// calculate equatorial coordinates (used by Slew command, takes Alt/Az -> moves telescope)
fbHor2Eq(alt := fElevation, 
		az := fAzimuth,
		jd := fJd+fTimeOffset,
		lat := telescopeConfig.latitude,
		lon := telescopeConfig.longitude,
		altitude := telescopeConfig.altitude,
		alt_is_observed := FALSE,
		ra => fRightAscensionCalc,
		dec => fDeclinationCalc,
		ha => fHourAngleCalc);		
// caluclate pointing offsets
fbPointingForward(
	HourAngle	:= fHourAngleApparent,
	Declination	:= fDeclinationApparent,
	Latitude	:= telescopeConfig.latitude,
	HourAngle_correction => fHourAnglePointingOffset,
	Declination_correction => fDeclinationPointingOffset,
	HourAngle_velocity => fHourAngleVelocity,
	Declination_velocity => fDeclinationVelocity,
);
(*--------------------------------------------------------------*)
// get current coordinates (of motors)
fDeclinationCurrent := fbDeclination.ActualPosition ;
fHourAngleCurrent := fbHourAngle.ActualPosition ;
// calculte pointing inversion
fbPointingInversion(
	HourAngle:= fHourAngleCurrent,
	Declination:= fDeclinationCurrent,
	Latitude:=telescopeConfig.latitude,
	HourAngle_correction => fHourAngleInversionOffsetCalc,
	Declination_correction => fDeclinationInversionOffsetCalc,
	bValid => bPointingInversionValid
);
// near the horizon the inversion is chaotic and does not converge (see FB_PointingModelInversion);
// keep reporting the last trustworthy correction rather than whatever garbage it would return
IF bPointingInversionValid THEN
	fHourAngleInversionOffset := fHourAngleInversionOffsetCalc;
	fDeclinationInversionOffset := fDeclinationInversionOffsetCalc;
END_IF
(*--------------------------------------------------------------*)
// transform from apparent to icrs

//current
fbHaDec2RaDec(
	ha := fHourAngleCurrent,
	dec := fDeclinationCurrent,
	jd := fJd+fTimeOffset,
	lon := telescopeConfig.longitude,
	ra_out => fRightAscensionCurrentICRS,
	dec_out => fDeclinationCurrentICRS);
//current corrected
fbHaDec2RaDec(
	ha := fHourAngleCurrent - fHourAngleInversionOffset - F_HourAngleOffsetOnAxis(fHourAngleOffset, fDeclinationApparent),
	dec := fDeclinationCurrent - fDeclinationInversionOffset- fDeclinationOffset,
	jd := fJd+fTimeOffset,
	lon := telescopeConfig.longitude,
	ra_out => fRightAscensionCurrentICRScorr,
	dec_out => fDeclinationCurrentICRScorr);
(*--------------------------------------------------------------*)
// to ALT AZ
fbEq2Hor(
	ra := fRightAscensionCurrentICRS,
	dec := fDeclinationCurrentICRS,
	lon := telescopeConfig.longitude,
	lat := telescopeConfig.latitude,
	altitude := telescopeConfig.altitude,
	refract_to_observed := FALSE,
	JD := fJd + fTimeOffset,
	alt => fElevationCurrent,
	az => fAzimuthCurrent);
	
fbEq2Hor(
	ra := fRightAscensionCurrentICRScorr,
	dec := fDeclinationCurrentICRScorr,
	lon := telescopeConfig.longitude,
	lat := telescopeConfig.latitude,
	altitude := telescopeConfig.altitude,
	refract_to_observed := FALSE,
	JD := fJd + fTimeOffset,
	alt => fElevationCurrentSky,
	az => fAzimuthCurrentSky);
END_METHOD

// Hook of the template body (BROTLib#25 step 5.4, S3: the body of this block is the template text, the differences are in these methods). Horizon and pole-zone guards, limit homes, target checks.
METHOD PROTECTED _Guards
// #161: while an axis is uncalibrated (e.g. after a PLC activation) its counter is meaningless, so the horizon and
// pole-zone stops must not act on it, otherwise the power-on sweep and the jog are stopped. Protection then is the NC
// software limits, the sweep's DistanceLimit and the operator.
bAxesCalibrated := fbHourAngle.Calibrated AND fbDeclination.Calibrated;
// losing the reference while enabled and not homing: stop instead of silently releasing the horizon protection
rtrigCalibLost(CLK := bAxesCalibrated);
IF rtrigCalibLost.Q AND bReady AND NOT bError AND NOT aAxis[1].bHoming AND NOT aAxis[2].bHoming THEN
	_AutoStop();
END_IF
// #166: a running power-on does not move a calibrated axis, but enabling it is not settled for a few scans and the mount
// is not ready before stage 100, so a mount inside a limit was stopped and the power-on aborted (any bStop aborts it).
// Skip the automatic stop only while the axes that matter stand still; stage 100 hands over to bGoHome. Any motion, a
// user stop or an error still stops.
bPowerOnHold := bPowerActive AND NOT bError;
bHaMoving := aAxis[1].bInMotion OR aAxis[1].bInRamp OR aAxis[1].bHoming;
bDecMoving := aAxis[2].bInMotion OR aAxis[2].bInRamp OR aAxis[2].bHoming;
// If the Telescope dips under the fHorizon (e.g. while tracking, stop and gohome)
// (also gated on fPointingSafeAltitude so tracking never lingers in the pointing model's chaotic zone)
// #84: a park requested in a limit homes out of it first and then parks. The stop conditions are unchanged.
IF NOT bGoHomeActive THEN
	bLimitHome := FALSE;
END_IF
IF NOT bParkActive THEN
	bParkAfterHome := FALSE;
	bParkHomeDone := FALSE;
	bParkForceInPlace := FALSE;
END_IF
bInHorizonLimit := bAxesCalibrated AND fElevationCurrent < MAX(fHorizon+0.2, fPointingSafeAltitude);
bInPoleLimit := (fbDeclination.Calibrated AND fDeclinationCurrent > (90.0 - fPoleZone)) OR (bAxesCalibrated AND bTrackActive AND (fDeclinationApparent + fDeclinationOffset + fDeclinationPointingOffset > (90.0 - fPoleZone)));
IF bInHorizonLimit THEN
	IF NOT bSettled AND NOT bGoHomeActive AND NOT (bPowerOnHold AND NOT bHaMoving AND NOT bDecMoving) THEN
		_AutoStop();
	ELSIF bReady AND NOT bError AND NOT bParkHomeDone THEN	// #82: only when the home can run; the power-on homes (stage 100)
		bGoHomeActive := TRUE;
		bLimitHome := TRUE;		// #84: also when bGoHome was set already (Home(), power-on stage 100)
	END_IF
END_IF
// If the Telescope goes into the forbidden polezone (e.g. while tracking, stop and gohome)
IF bInPoleLimit THEN
	IF NOT bSettled AND NOT bGoHomeActive AND NOT (bPowerOnHold AND NOT bDecMoving) THEN
		_AutoStop();
	ELSIF bReady AND NOT bError AND NOT bParkHomeDone THEN	// #82: only when the home can run; the power-on homes (stage 100)
		bGoHomeActive := TRUE;
		bLimitHome := TRUE;		// #84
	END_IF
END_IF
//----------------------------------------------------------------------------------------------
// if the given coordinates to goto/slew are under the horizon
// (also rejects targets below fPointingSafeAltitude, where the pointing model's inversion is chaotic -- see FB_PointingModelInversion)
IF (bGotoActive AND (fElevationCalc < MAX(fHorizon + 1.0, fPointingSafeAltitude))) OR (bSlewActive AND (fElevation < MAX(fHorizon, fPointingSafeAltitude))) THEN
	// trigger event
	rtrigHorizonError(CLK:=TRUE);
	// reset input coords to parking position (always over horizon to stop bHorizonError from occuring)
	fDeclination := telescopeConfig.declinationPark;
	fbHaDec2RaDec(	jd := fJd +fTimeOffset,
					ha := telescopeConfig.houranglePark,
					dec := telescopeConfig.declinationPark,
					lon := telescopeConfig.longitude,
					ra_out => fRightAscension);
	// reset elevation values to abitrarry value over horizon, will get overwritten down the line
	fElevationCalc := 20.0;
	fElevation := 20.0;
	// stop telescope
	_AutoStop();
ELSE
	// reset event trigger
	rtrigHorizonError(CLK:=FALSE);
END_IF

// if the given coordinates to goto/slew are in the PoleZone
IF (bGotoActive AND (fDeclinationApparent > (90.0 - fPoleZone))) OR (bSlewActive AND (fDeclinationCalc  > (90.0 - fPoleZone))) THEN
	// trigger event
	rtrigPoleError(CLK:=TRUE);
	// reset input coords to parking position (always over horizon to stop bHorizonError from occuring)
	fDeclination := telescopeConfig.declinationPark;
	fbHaDec2RaDec(	jd := fJd +fTimeOffset,
					ha := telescopeConfig.houranglePark,
					dec := telescopeConfig.declinationPark,
					lon := telescopeConfig.longitude,
					ra_out => fRightAscension);
	// reset elevation values to abitrarry value over horizon, will get overwritten down the line
	fElevationCalc := 20.0;
	fElevation := 20.0;
	// stop telescope
	_AutoStop();

ELSE
	// reset event trigger
	rtrigPoleError(CLK:=FALSE);
END_IF
END_METHOD

// Hook of the template body (BROTLib#25 step 5.4, S3: the body of this block is the template text, the differences are in these methods). Power-on warning, idle park, state-machine timeouts, pending home and park.
METHOD PROTECTED _Timers
tpPowerOnWarning(IN := bPowerActive OR (NOT fbHourAngle.bEnable), PT := T#250MS);

tonPowerTimeout(IN := TCS_command = E_TCSCommand.no_command AND NOT bIsParked, PT := T#12H, nDivisor := nTimeDivisor);
// MONETcommon#17: state-machine timeouts, checked in _GotoTelescope/_HomeTelescope/_SlewTelescope
// #75: count only while the command is the one being run (TCS_command is last scan's dispatch) and without an error.
// Counting from the request, a command that never started (not ready, preempted) fired the timeout in the next
// stop/park/reset after 600 s and latched an error, and with the horizon/pole auto-home setting bGoHome again every
// scan the timer never dropped, so no reset cleared it.
tonGotoTimeout(IN := bGotoActive AND TCS_command = E_TCSCommand.goto AND NOT bError, PT := T#600S, nDivisor := nTimeDivisor);
tonHomeTimeout(IN := bGoHomeActive AND TCS_command = E_TCSCommand.gohome AND NOT bError, PT := T#600S, nDivisor := nTimeDivisor);
tonSlewTimeout(IN := bSlewActive AND TCS_command = E_TCSCommand.slew AND NOT bError, PT := T#600S, nDivisor := nTimeDivisor);
tonParkTimeout(IN := bParkActive AND TCS_command = E_TCSCommand.park AND NOT bError, PT := T#600S, nDivisor := nTimeDivisor);
// #75: a Home() that never starts (axes off, telescope not ready) left bGoHome set for good, swallowing Track() and
// Slew(). Drop it after 2 min, with a log line, without an error. Not at once: the home that the power-on requests in
// stage 100 can wait a few scans for bReady, and a stop from slew speed takes about 4 s. Not during a power-on.
tonHomePending(IN := bGoHomeActive AND TCS_command <> E_TCSCommand.gohome AND NOT bPowerActive AND NOT bError, PT := T#2M, nDivisor := nTimeDivisor);
IF tonHomePending.Q THEN
    fbStartup.MarkAbortedIfInitializing();
	bGoHomeActive := FALSE;
	// #108: say what was pending. "Not ready, power on" was also logged when a stop before the home had not finished.
	fbHomeDrop(bReady := bReady, bStopPending := TCS_command = E_TCSCommand.stop OR NOT bSettled);
	sHomeEnd := fbHomeDrop.sEnd;
	sHomeDropWhy := fbHomeDrop.sWhy;
	bHomeCancelled := TRUE;
END_IF
// #197: a park that is requested but not started (not dispatched, not in the axes-off path, no stop or home running)
// waited without a timeout: tonParkTimeout counts only a running park (#75). After 2 min: say why and park in place.
tonParkPending(IN := bParkActive AND TCS_command <> E_TCSCommand.park AND TCS_command <> E_TCSCommand.gohome
	AND NOT bMoveAbortPending AND NOT bError AND NOT bEstopTriggered AND NOT bParkForceInPlace, PT := T#2M, nDivisor := nTimeDivisor);
IF tonParkPending.Q THEN
	bParkForceInPlace := TRUE;
	fbHomeDrop(bReady := bReady, bStopPending := TCS_command = E_TCSCommand.stop OR NOT bSettled);
	TCSparkErrorEvent.OnMessage := CONCAT(CONCAT('Park did not start within 2 min (', fbHomeDrop.sWhy), '): parking in place with the axes off.');
	bParkInError := TRUE;
END_IF
IF tonPowerTimeout.Q AND NOT bIsParked THEN
	bParkActive := TRUE;
	// #83: fire once. With the axes off or in error the park does not set bIsParked, so Q stayed TRUE and bPark was
	// set again every scan (dropping Track/Goto/Slew/Home, re-commanding the dome). The timer counts again from now.
	tonPowerTimeout(IN := FALSE);
END_IF
END_METHOD

// Hook of the template body (BROTLib#25 step 5.4, S3: the body of this block is the template text, the differences are in these methods). The replacement gets its own timeout.
METHOD PROTECTED _RestartMoveTimeout
VAR_INPUT
	eKeep	: E_TCSCommand;
END_VAR
CASE eKeep OF
	E_TCSCommand.gohome:	tonHomeTimeout(IN := FALSE, PT := T#600S, nDivisor := nTimeDivisor);
	E_TCSCommand.goto:		tonGotoTimeout(IN := FALSE, PT := T#600S, nDivisor := nTimeDivisor);
	E_TCSCommand.slew:		tonSlewTimeout(IN := FALSE, PT := T#600S, nDivisor := nTimeDivisor);
END_CASE
END_METHOD

// Hook of the template body (BROTLib#25 step 5.4, S3: the body of this block is the template text, the differences are in these methods). The automatic parks.
METHOD PROTECTED _ParkRequests
// BROTLib#25 step 4.4d (decided by Tim 2026-11-09: MONETcommon wins): a new hardware error (hour angle, declination or focus; not a
// software or cabinet error) while not parked and without E-stop starts the park by itself, like MONETcommon#86. The park branch
// below does what is safe without the mount (the axes are disabled by the error): covers close, dome parks, focus off; the mount
// is not moved and bIsParked is not set until the covers are closed and the dome is parked. A running power-on is aborted by
// the park (#109). Edge only: a still present error does not start it again.
bErrorParkStarted := BROTLib.F_ErrorParkRequest(
	bHwError := fbHourAngle.Error OR fbDeclination.Error OR (fbFocus <> 0 AND_THEN fbFocus.Error),
	bHwErrorLast := bHwErrorLast,
	bIsParked := bIsParked,
	bEstop := bEstopTriggered);
bHwErrorLast := fbHourAngle.Error OR fbDeclination.Error OR (fbFocus <> 0 AND_THEN fbFocus.Error);
IF bErrorParkStarted THEN
	Park();
END_IF
END_METHOD

// Hook of the template body (BROTLib#25 step 5.4, S3: the body of this block is the template text, the differences are in these methods). TRUE: the pending park waits. The gate (no stop, no power-on, no abort stop) is in the body.
METHOD PROTECTED _ParkPreStep : BOOL
_ParkPreStep := FALSE;
bTrackActive := FALSE;
IF bError OR bEstopTriggered OR (TCS_command <> E_TCSCommand.park AND NOT fbHourAngle.Enable AND NOT fbDeclination.Enable) THEN
	_ParkInPlace();
	_ParkPreStep := TRUE;
ELSIF (NOT bIsPowered OR bParkForceInPlace) AND TCS_command <> E_TCSCommand.park THEN
	// #197: no completed power-on (aborted by this park, or stopped in stage 40 or later) but an axis is on: the park can
	// never be dispatched. Switch the axes off once they are at rest, then the axes-off park parks in place.
	// TCS_command must not stay on poweron: _PowerOn and its 12 h timeout would stay selected.
	fbSweepStop.ArmAll();
	TCS_command := E_TCSCommand.no_command;
	_ParkPreStep := TRUE;
ELSIF bGoHomeActive AND bLimitHome THEN
	// #84: a park in a limit: the home out of the limit runs first (the arbiter dispatches it), the park follows (bParkHomeDone)
	IF NOT bParkAfterHome THEN
		bParkAfterHome := TRUE;
		bParkHomeFirst := TRUE;
	END_IF
	_ParkPreStep := TRUE;
ELSIF NOT (bReady AND NOT bBusy) THEN
	_ParkPreStep := TRUE;
END_IF
END_METHOD

// Hook of the template body (BROTLib#25 step 5.4, S3: the body of this block is the template text, the differences are in these methods). The arbiter input bEmergencyPark.
METHOD PROTECTED _EmergencyPark : BOOL
_EmergencyPark := FALSE;
END_METHOD

// Hook of the template body (BROTLib#25 step 5.4, S3: the body of this block is the template text, the differences are in these methods). The arbiter input bStopped: at rest and no stop transaction running.
METHOD PROTECTED _AtRest : BOOL
_AtRest := bSettled;	// IAG50cm: at rest and no stop transaction running
END_METHOD

// Hook of the template body (BROTLib#25 step 5.4, S3: the body of this block is the template text, the differences are in these methods). The arbiter interrupts the power-on.
METHOD PROTECTED _InterruptPower
IF _PowerOnStage() >= 40 THEN	// abort path: bPowerActive FALSE, startup marked aborted, stage 0; returns the stage it was in
	IF fbArbiter.bPowerAbortedByPark THEN
		// #197: the axes are on and may be sweeping: stop them. The park then switches them off (nothing else can: bReady
		// needs the completed power-on) and parks in place.
		fbSweepStop.ArmAll();
	ELSE
		fbSweepStop.Arm();		// #113: stopped in the calibration sweep (stage 40 and later)
	END_IF
	fbHourAngle.bStopSweep := TRUE;		// #198: no new sweep step after this stop, also before the sweep has started
	fbDeclination.bStopSweep := TRUE;
END_IF
END_METHOD

// Hook of the template body (BROTLib#25 step 5.4, S3: the body of this block is the template text, the differences are in these methods). The arbiter interrupts the park.
METHOD PROTECTED _InterruptPark
IF bWasPark THEN
	sParkEnd := 'cancelled by stop';
	fbSweepStop.Cancel();		// #197: the park is gone, the axes stay as they are
END_IF
_DoPark();
END_METHOD

// Hook of the template body (BROTLib#25 step 5.4, S3: the body of this block is the template text, the differences are in these methods). The arbiter interrupts the goto.
METHOD PROTECTED _InterruptGoto
_DoGoto();
END_METHOD

// Hook of the template body (BROTLib#25 step 5.4, S3: the body of this block is the template text, the differences are in these methods). The arbiter interrupts the slew.
METHOD PROTECTED _InterruptSlew
_DoSlew();
END_METHOD

// Hook of the template body (BROTLib#25 step 5.4, S3: the body of this block is the template text, the differences are in these methods). The arbiter interrupts the home.
METHOD PROTECTED _InterruptGoHome
IF bWasGoHome THEN
	IF bStopActive THEN
		sHomeEnd := 'cancelled by stop';	// #84: also the home that a park waited for
	ELSE
		sHomeEnd := 'cancelled by park';
	END_IF
END_IF
_DoGoHome();
END_METHOD

// Hook of the template body (BROTLib#25 step 5.4, S3: the body of this block is the template text, the differences are in these methods). After the arbiter has been applied.
METHOD PROTECTED _AfterArbiter
// #196: the axes are off, there is nothing to stop; the covers have no stop command and the park goes on
IF bStopActive AND bSafeParked AND NOT bWasPark AND NOT bWasPower AND NOT bWasMove AND NOT bWasGoHome THEN
	bStopIgnored := TRUE;
END_IF
END_METHOD

// Hook of the template body (BROTLib#25 step 5.4, S3: the body of this block is the template text, the differences are in these methods). Idle: the axis commands are dropped.
METHOD PROTECTED _DropAxisCommands
	fbHourAngle.MoveAxis := FALSE;
	fbDeclination.MoveAxis := FALSE;
	fbHourAngle.bTracking := FALSE;
	fbDeclination.bTracking := FALSE;
END_METHOD

// Hook of the template body (BROTLib#25 step 5.4, S3: the body of this block is the template text, the differences are in these methods). TCS_command changed.
METHOD PROTECTED _OnCommandChanged
// #108: a stop transaction starts here and lasts as long as TCS_command stays stop (also through the wait of a
// gohome that preempted a track): each axis gets one stop in it
IF TCS_command = E_TCSCommand.stop THEN
	fbStopTx.Begin();
END_IF
END_METHOD

// Calls the stage machine of the power-on; returns the stage it was in (>= 40: the sweep stop of the power-on runs).
METHOD PRIVATE _PowerOnStage : USINT
_PowerOnStage := _PowerOn();
END_METHOD

// Hook of the template body (BROTLib#25 step 5.4). Calls the stage machine of the power-on.
METHOD PROTECTED _DoPowerOn
_PowerOnStage();
END_METHOD

// Hook of the template body (BROTLib#25 step 5.4, S3: the body of this block is the template text, the differences are in these methods). Calls the stage machine.
METHOD PROTECTED _DoPark
_ParkTelescope();
END_METHOD

// Hook of the template body (BROTLib#25 step 5.4, S3: the body of this block is the template text, the differences are in these methods). Calls the stage machine.
METHOD PROTECTED _DoGoHome
_HomeTelescope();
END_METHOD

// Hook of the template body (BROTLib#25 step 5.4, S3: the body of this block is the template text, the differences are in these methods). Calls the stage machine.
METHOD PROTECTED _DoGoto
_GotoTelescope();
END_METHOD

// Hook of the template body (BROTLib#25 step 5.4, S3: the body of this block is the template text, the differences are in these methods). Calls the stage machine.
METHOD PROTECTED _DoSlew
_SlewTelescope();
END_METHOD

// Hook of the template body (BROTLib#25 step 5.4, S3: the body of this block is the template text, the differences are in these methods). Calls the stage machine.
METHOD PROTECTED _DoTrack
_TrackTelescope();
END_METHOD

// Hook of the template body (BROTLib#25 step 5.4, S3: the body of this block is the template text, the differences are in these methods). Calls the stage machine.
METHOD PROTECTED _DoStop
_StopTelescope();
END_METHOD

// Hook of the template body (BROTLib#25 step 5.4, S3: the body of this block is the template text, the differences are in these methods). The timeout of a command.
METHOD PROTECTED _CommandTimeout : TIME
VAR_INPUT
	eCommand	: E_TCSCommand;
END_VAR
CASE eCommand OF
	E_TCSCommand.poweron:	_CommandTimeout := T#12H;
	E_TCSCommand.stop:		_CommandTimeout := T#30S;	// #40: a stop from slew speed takes about 4 s, a preempting stop can follow a long move
	E_TCSCommand.track:		_CommandTimeout := T#12H;
ELSE
	_CommandTimeout := T#2M;
END_CASE
END_METHOD

// Hook of the template body (BROTLib#25 step 5.4, S3: the body of this block is the template text, the differences are in these methods). After the dispatch.
METHOD PROTECTED _AfterDispatch
// nothing
END_METHOD

// Hook of the template body (BROTLib#25 step 5.4, S3: the body of this block is the template text, the differences are in these methods). Motion, stop transaction, sweep stop, readiness and the in-place park status.
METHOD PROTECTED _UpdateStatus
(* STATUS BOOLS*)
bSliding := NOT bTracking AND (aAxis[1].bInMotion OR aAxis[1].bInRamp OR
			aAxis[2].bInMotion OR aAxis[2].bInRamp );

// signal must be stable for 1s
tonTrackingDelay(in := aAxis[1].bTracking AND
			aAxis[2].bTracking ,PT :=T#1000MS, Q => bTracking);

// #92: a move that was commanded (MoveAxis -> MoveTo) is reported by the NC a few cycles later; until then the axis
// reports StandStill. A stop in that window saw bStopped, so bStop was cleared after one scan, the stop only dropped
// MoveAxis (which does not cancel a move that has started) and no axis stop was sent: the move ran to its end (T18.4,
// park, Dec). The axis is not at rest while its move is on the way; the stop then lasts until the axis moves and gets
// its axis stop from the stop transaction.
rtHaMove(CLK := fbHourAngle.MoveAxis);
rtDecMove(CLK := fbDeclination.MoveAxis);
IF rtHaMove.Q THEN
	bHaMovePending := TRUE;
END_IF
IF rtDecMove.Q THEN
	bDecMovePending := TRUE;
END_IF
IF aAxis[1].bInMotion OR aAxis[1].bInRamp OR aAxis[1].bHoming OR fbHourAngle.MoveDone OR bError OR NOT fbHourAngle.bEnable THEN
	bHaMovePending := FALSE;
END_IF
IF aAxis[2].bInMotion OR aAxis[2].bInRamp OR aAxis[2].bHoming OR fbDeclination.MoveDone OR bError OR NOT fbDeclination.bEnable THEN
	bDecMovePending := FALSE;
END_IF
tonHaMovePending(IN := bHaMovePending, PT := T#1S);
tonDecMovePending(IN := bDecMovePending, PT := T#1S);
IF tonHaMovePending.Q THEN
	bHaMovePending := FALSE;
END_IF
IF tonDecMovePending.Q THEN
	bDecMovePending := FALSE;
END_IF

// #198: a pause of the calibration sweep reports StandStill, but FB_LatchHome is still in its sequence (or about to start
// it): the axis is not at rest. A stop in a pause saw bStopped, ran for one scan and sent no axis stop.
bStopped :=  (NOT fbHourAngle.bEnable OR (aAxis[1].bStandStill AND NOT fbHourAngle.bSweepActive)) AND
			(NOT fbDeclination.bEnable OR (aAxis[2].bStandStill AND NOT fbDeclination.bSweepActive)) AND
			NOT bHaMovePending AND NOT bDecMovePending;

// #98: bStopped is TRUE for one scan at the start of every stop, before MC_Stop has taken hold (StandStill is still
// TRUE), and a home commanded while MC_Stop locks the axis (StateDWord bit 29) fails with 17135. A stop transaction
// is settled when every axis that was sent a stop reported Done and no axis has been locked for 3 scans.
IF bResetActive OR bError OR bEstopTriggered THEN
	fbStopTx.Cancel();
	fbSweepStop.Cancel();
END_IF
_SetStopTxInputs();
fbStopTx.Monitor();
bSettled := bStopped AND NOT fbStopTx.bActive;

// #120: a stop transaction that is not settled 30 s after it began (an axis never reported Done) no longer waits for the
// Done: it settles as soon as the telescope is at rest. The stop is not sent again. Clear StopAxis of the axes without a
// Done so that the next stop gives a rising edge (FB_AxisControl.StopAxis) and the home hold does not see a stale stop.
IF fbStopTx.bTimedOut THEN
	IF fbStopTx.abNoDone[1] AND fbStopTx.abNoDone[2] THEN
		sStopNoDone := 'HA and Dec';
	ELSIF fbStopTx.abNoDone[1] THEN
		sStopNoDone := 'HA';
	ELSE
		sStopNoDone := 'Dec';
	END_IF
	IF NOT fbStopTx.bActive THEN
		TCSstopTimeoutEvent.OnMessage := CONCAT(CONCAT('STOP: no stop Done from ', sStopNoDone), ' within 30 s; telescope at rest, stop released.');
	ELSIF NOT bStopped THEN
		TCSstopTimeoutEvent.OnMessage := CONCAT(CONCAT('STOP: no stop Done from ', sStopNoDone), ' within 30 s; axes still moving, released when at rest.');
	ELSE
		TCSstopTimeoutEvent.OnMessage := CONCAT(CONCAT('STOP: no stop Done from ', sStopNoDone), ' within 30 s; axis locked (stop active) or homing, released when it ends.');
	END_IF
	bStopTimeoutLog := TRUE;
ELSIF fbStopTx.bForced THEN
	TCSstopTimeoutEvent.OnMessage := 'STOP released: at rest without a stop Done from an axis (30 s timeout).';
	bStopTimeoutLog := TRUE;
END_IF
IF fbStopTx.bForced THEN
	IF fbStopTx.abNoDone[1] THEN
		fbHourAngle.StopAxis := FALSE;
	END_IF
	IF fbStopTx.abNoDone[2] THEN
		fbDeclination.StopAxis := FALSE;
	END_IF
END_IF

// #113: a stop in the calibration sweep leaves the axes enabled and uncalibrated; once the stop has settled and the
// homing is aborted, switch the uncalibrated axes off (the next power-on starts the sweep again), READY_STATE -2
IF bPowerActive THEN
	fbSweepStop.Cancel();
END_IF
fbSweepStop(bSettled := bSettled,
			bHaCalibrated := fbHourAngle.bCalibrated, bDecCalibrated := fbDeclination.bCalibrated,
			bHaHoming := fbHourAngle.fbLatchHome.Busy, bDecHoming := fbDeclination.fbLatchHome.Busy,
			bOtherBusy := fbFocus <> 0 AND_THEN fbFocus.Busy);
IF fbSweepStop.bDisableHa THEN
	fbHourAngle.Enable := FALSE;
END_IF
IF fbSweepStop.bDisableDec THEN
	fbDeclination.Enable := FALSE;
END_IF
			
bHomed := fbHourAngle.bCalibrated AND fbDeclination.bCalibrated AND (fbFocus <> 0 AND_THEN fbFocus.Calibrated);
			
bReady := bHomed AND 
	bIsPowered AND 
	fbHourAngle.bEnable AND
	fbDeclination.bEnable AND
	(fbFocus <> 0 AND_THEN fbFocus.Enable) AND
    NOT bError;

bBusy := aAxis[1].bBusy OR aAxis[2].bBusy OR (fbFocus <> 0 AND_THEN fbFocus.Busy);
//----------------------------------------------------------------------------------------------
(* STATUS STATES*)
// Public completion is latched only by the final startup stage, never by mechanical bReady alone.
// #110: the covered state ends with a power-on, an error or an E-stop.
IF bSafeParked AND (bPowerActive OR bError OR bEstopTriggered) THEN
	// #200: every exit of the in-place park has an end line
	IF bEstopTriggered THEN
		sParkInPlaceEnd := 'aborted: E-stop pressed, the covers and the dome cannot move. Release it, reset, then park again.';
		nParkInPlaceLevel := ADSLOG_MSGTYPE_WARN;
	ELSIF bError THEN
		IF fbCovers.Closed THEN
			sParkInPlaceEnd := 'aborted by an error: covers closed, the mount was not moved. Reset, then park again.';
		ELSE
			sParkInPlaceEnd := 'aborted by an error: covers closing, the mount was not moved. Reset, then park again.';
		END_IF
		nParkInPlaceLevel := ADSLOG_MSGTYPE_WARN;
	ELSE
		sParkInPlaceEnd := 'cancelled by power-on';
		nParkInPlaceLevel := ADSLOG_MSGTYPE_HINT;
	END_IF
	bParkInPlaceDone := TRUE;
END_IF
IF bPowerActive OR bError OR bEstopTriggered THEN
    bSafeParked := FALSE;
END_IF
// #187: an axes-off park (power-on aborted by a park, park after a stopped power-on) ends parked, like a park of MONET:
// bIsParked means covers closed and dome parked with the axes off, bParkedInPlace says the mount was not moved.
// Without it bIsParked stayed FALSE, and the 12 h idle park fired again every 12 h.
tonParkInPlace(IN := bSafeParked AND NOT bIsParked, PT := T#120S, nDivisor := nTimeDivisor);
IF bSafeParked AND fbCovers.Closed AND fbDome.Parked THEN
	IF NOT bIsParked OR bParkInPlaceOpen THEN
		bIsParked := TRUE;
		bParkedInPlace := TRUE;
		sParkInPlaceEnd := 'completed in place: covers closed, dome parked, the mount stays where it stood (#187)';
		nParkInPlaceLevel := ADSLOG_MSGTYPE_HINT;
		bParkInPlaceDone := TRUE;
	END_IF
	bIsPowered := FALSE;
	bSafeParked := FALSE;
ELSIF bSafeParked AND (tonParkInPlace.Q OR fbDome.Error) THEN
	// give up: not 0.3 for ever. The park start line said what was requested; this is the end line (#200).
	bSafeParked := FALSE;
	sParkInPlaceEnd := 'aborted: the covers did not close or the dome did not park within 120 s, or the dome is in error.';
	nParkInPlaceLevel := ADSLOG_MSGTYPE_WARN;
	bParkInPlaceDone := TRUE;
END_IF
END_METHOD

// Hook of the template body (BROTLib#25 step 5.4, S3: the body of this block is the template text, the differences are in these methods). The Parking input of the READY_STATE.
METHOD PROTECTED _ReadyStateParking : BOOL
_ReadyStateParking := (bParkActive OR bSafeParked) AND NOT bPowerActive;
END_METHOD

// Hook of the template body (BROTLib#25 step 5.4, S3: the body of this block is the template text, the differences are in these methods). The slewing flag of the motion state.
METHOD PROTECTED _IsSlewing : BOOL
_IsSlewing := bSliding;
END_METHOD

// Hook of the template body (BROTLib#25 step 5.4, S3: the body of this block is the template text, the differences are in these methods). The stop transaction has settled.
METHOD PROTECTED _StopSettled : BOOL
_StopSettled := bSettled;
END_METHOD

// Hook of the template body (BROTLib#25 step 5.4, S3: the body of this block is the template text, the differences are in these methods). The abort stop has been released.
METHOD PROTECTED _OnAbortStopReleased
// nothing
END_METHOD

// Hook of the template body (BROTLib#25 step 5.4, S3: the body of this block is the template text, the differences are in these methods). The reset is released.
METHOD PROTECTED _ReleaseReset
// unset the RESET command when no Error is present
IF NOT bError THEN
	bResetActive := FALSE;
END_IF
END_METHOD

// Hook of the template body (BROTLib#25 step 5.4, S3: the body of this block is the template text, the differences are in these methods). End of the scan: the drives are cut on an E-stop.
METHOD PROTECTED _SafeStateEndOfScan
IF bEstopTriggered THEN
	fbHourAngle.Enable := FALSE;
	fbDeclination.Enable := FALSE;
END_IF
END_METHOD

// Hook of the template body (BROTLib#25 step 5.4, S3: the body of this block is the template text, the differences are in these methods). The period of the telemetry.
METHOD PROTECTED _TelemetryPeriod : TIME
IF bSliding OR bTrackActive OR bTracking THEN
	_TelemetryPeriod := T#1000MS;	// during movement every second
ELSE
	_TelemetryPeriod := T#5000MS;	// otherwise every five seconds
END_IF
END_METHOD

// Hook of the template body (BROTLib#25 step 5.4, S3: the body of this block is the template text, the differences are in these methods). Sends the telemetry.
METHOD PROTECTED _SendTelemetry : BOOL
THIS^._SendTelemetryEquitorial();
END_METHOD

// Hook of the template body (BROTLib#25 step 5.4, S3: the body of this block is the template text, the differences are in these methods). End of the scan.
METHOD PROTECTED _EndOfScan
IF NOT bGoHomeActive AND TCS_command <> E_TCSCommand.gohome THEN
	bHomeByCommand := FALSE;	// the commanded home is over
END_IF
END_METHOD

// plan step 3.4: the event function blocks at the end of the body (ADS log and MQTT log), moved unchanged; called at the end of the body.
METHOD PROTECTED _LogEvents
VAR_INPUT
END_VAR
(* Event function blocks start here. *)
TCSpowerEvent(	Trigger := bPowerFailure, 
				Level := ADSLOG_MSGTYPE_ERROR,
				FormatString := 'power %s',
				//OnMessage := 'Failure',
				OffMessage := 'OK', 
				Comm := fbComm);

TCSgohomeEvent.OffMessage := sHomeEnd;		// #75: "GOHOME completed" was also logged when the home was cancelled or timed out
TCSgohomeEvent(	Trigger := bGoHomeActive, 
				Level := ADSLOG_MSGTYPE_HINT,
				FormatString := 'GOHOME %s',
				OnMessage := 'commencing',
				Comm := fbComm);
sHomeEnd := 'completed';
// #197/#200: the in-place park that goes on from a logged park ends with the PARK end line, one per park
IF bParkInPlaceDone AND bParkInPlaceOpen THEN
	sParkEnd := sParkInPlaceEnd;
	TCSparkEvent.OffLevel := nParkInPlaceLevel;
	bParkInPlaceOpen := FALSE;
	bParkInPlaceDone := FALSE;
END_IF
TCSparkEvent.OffMessage := sParkEnd;		// #57: "PARK completed" was also logged when the park was cancelled
TCSparkEvent(	Trigger := bParkActive OR bParkInPlaceOpen,
				Level := ADSLOG_MSGTYPE_HINT,
				FormatString := 'PARK %s',
				OnMessage := 'commencing',
				Comm := fbComm);
TCSparkInPlaceEvent(	Trigger := bParkInPlaceDone,
				Level := nParkInPlaceLevel,
				FormatString := 'PARK %s',
				OnMessage := sParkInPlaceEnd,
				Comm := fbComm);
bParkInPlaceDone := FALSE;
bParkLogged := bParkActive;
sParkEnd := 'completed';
TCSparkEvent.OffLevel := ADSLOG_MSGTYPE_HINT;
TCSgotoEvent(	Trigger := bGotoActive, 
				Level := ADSLOG_MSGTYPE_HINT,
				FormatString := 'GOTO %s',
				OnMessage := 'commencing',
				OffMEssage := 'completed', 
				Comm := fbComm);
TCStrackEvent(	Trigger := bTrackActive, 
				Level := ADSLOG_MSGTYPE_HINT,
				FormatString := 'TRACK %s',
				OnMessage := 'commencing',
				OffMEssage := 'completed', 
				Comm := fbComm);
TCSstopEvent(	Trigger := bStopActive, 
				Level := ADSLOG_MSGTYPE_WARN,
				FormatString := 'STOP %s',
				OnMessage := 'commencing',
				OffMEssage := 'completed',
				OffLevel := ADSLOG_MSGTYPE_HINT, 
				Comm := fbComm);
TCSstopIgnoredEvent(	Trigger := bStopIgnored,
				Level := ADSLOG_MSGTYPE_WARN,
				FormatString := '%s',
				OnMessage := 'Stop ignored: the covers and the dome cannot be stopped, the in-place park continues.',
				Comm := fbComm);
bStopIgnored := FALSE;
TCStargetHorizonEvent(	Trigger := rtrigHorizonError.Q, 
				Level := ADSLOG_MSGTYPE_WARN,
				FormatString := '%s',
				OnMessage := 'Target below safe horizon, stopping telescope.',
				OffMEssage := '', 
				Comm := fbComm);
TCSaltitudeEvent(	Trigger := bAxesCalibrated AND fElevationCurrent<MAX(fHorizon+2.0, fPointingSafeAltitude+2.0),
				Level := ADSLOG_MSGTYPE_WARN,
				FormatString := '%s',
				OnMessage := 'Telescope below safe horizon, aboard and slew telescope to home position.',
				OffMEssage := '', 
				Comm := fbComm);
TCSnearPoleEvent(	Trigger := rtrigPoleError.Q, 
				Level := ADSLOG_MSGTYPE_WARN,
				FormatString := '%s',
				OnMessage := 'Target to close to the celestial pole, stopping telescope.',
				OffMEssage := '', 
				Comm := fbComm);			
TCSreadyEvent(	Trigger := bReady, 
				Level := ADSLOG_MSGTYPE_HINT,
				FormatString := '%s',
				OnMessage := 'IAG50cm startup finished', 
				Comm := fbComm);
TCSparkErrorEvent(	Trigger := bParkInError,
				Level := ADSLOG_MSGTYPE_WARN,
				FormatString := '%s',
				// OnMessage is set in the arbitration (texts built from sParkWhy); a literal here overwrote it (#57)
				Comm := fbComm);
bParkInError := FALSE;
TCShomeCancelEvent(	Trigger := bHomeCancelled,
				Level := ADSLOG_MSGTYPE_WARN,
				FormatString := '%s',
				OnMessage := CONCAT('Home request dropped: ', sHomeDropWhy),
				Comm := fbComm);
bHomeCancelled := FALSE;
TCSpowerBlockedEvent(	Trigger := bPowerBlocked,
				Level := ADSLOG_MSGTYPE_ERROR,
				FormatString := '%s',
				Comm := fbComm);
bPowerBlocked := FALSE;
TCSparkHomeEvent(	Trigger := bParkHomeFirst,
				Level := ADSLOG_MSGTYPE_HINT,
				FormatString := '%s',
				OnMessage := 'Park in the horizon/pole-zone limit: homing out of it first, then parking',
				Comm := fbComm);
bParkHomeFirst := FALSE;
TCSpowerParkEvent(	Trigger := bPowerAbortedByPark,
				Level := ADSLOG_MSGTYPE_WARN,
				FormatString := '%s',
				OnMessage := 'Power-on aborted by park',
				Comm := fbComm);
bPowerAbortedByPark := FALSE;
TCSinitRefusedEvent(	Trigger := bInitRefused,
				Level := ADSLOG_MSGTYPE_WARN,
				FormatString := 'power-on ignored: %s',
				OnMessage := sInitRefusedReason,
				Comm := fbComm);
bInitRefused := FALSE;
// every rejection is logged (ADS log and MQTT log topic); an identical one repeated within 2 s once, all are counted. The event is
// re-armed with FALSE first so that rejections in consecutive scans each give a rising edge (as MONETcommon).
tonRejectRepeat(IN := TRUE, PT := T#2S);
RejectEvent(Trigger := FALSE, Comm := fbComm);
IF bCommandRejected THEN
	IF tonRejectRepeat.Q OR eLastRejectedCommand <> eLoggedCommand OR eLastRejectReason <> eLoggedReason THEN
		sRejectMessage := CONCAT(CONCAT(BROTLib.F_TCSCommandText(eLastRejectedCommand), ' rejected: '),
			BROTLib.F_CommandRejectText(eLastRejectReason));
		RejectEvent(Trigger := TRUE, Level := ADSLOG_MSGTYPE_WARN, FormatString := '%s',
			OnMessage := sRejectMessage, Comm := fbComm);
		eLoggedCommand := eLastRejectedCommand;
		eLoggedReason := eLastRejectReason;
		tonRejectRepeat(IN := FALSE);
	END_IF
	bCommandRejected := FALSE;
END_IF
TCSstopTimeoutEvent(	Trigger := bStopTimeoutLog,
				Level := ADSLOG_MSGTYPE_WARN,
				FormatString := '%s',
				Comm := fbComm);
bStopTimeoutLog := FALSE;
TCSsoftErrorEvent(	Trigger := bSoftwareError,
				Level := ADSLOG_MSGTYPE_ERROR,
				FormatString := 'Command timeout error %s',	// 16 goto, 32 park, 48 gohome, 64 slew (16#10, 16#20, 16#30, 16#40)
				OnMessage := UDINT_TO_STRING(nSoftwareErrorID),
				OffMessage := 'reset',
				Comm := fbComm);
TCSCTOEvent(	Trigger := tonCommandTimeout.Q,
				Level := ADSLOG_MSGTYPE_WARN,
				FormatString := 'A timeout occured during %s command!',
				Comm := fbComm);
END_METHOD

// The state BROTLib.F_CommandAcceptance decides on. eExcludeOwn leaves the own request out of bMoveActive. bMoveAbortPending stands in for
// bMoveAbortPending until the abort stop (command model step 3A).
METHOD PRIVATE _CommandState : BROTLib.ST_CommandState
VAR_INPUT
	eExcludeOwn	: E_TCSCommand;
END_VAR
_CommandState.bEstop		:= bEstopTriggered;
_CommandState.bError		:= bError;
_CommandState.bClockValid	:= fbTime.bValid;
_CommandState.bStop			:= bStopActive;
_CommandState.bPowering		:= bPowerActive OR fbStartup.Initializing;
_CommandState.bParkPending	:= bParkActive OR bParkAfterStop;
_CommandState.bIsParked		:= bIsParked;
_CommandState.bReady		:= bReady;
_CommandState.bGoHomeActive	:= bHomeByCommand AND ((bGoHomeActive AND eExcludeOwn <> E_TCSCommand.gohome) OR TCS_command = E_TCSCommand.gohome);
_CommandState.bMoveActive	:= (bGotoActive AND eExcludeOwn <> E_TCSCommand.goto) OR
	(bSlewActive AND eExcludeOwn <> E_TCSCommand.slew) OR
	(bTrackActive AND eExcludeOwn <> E_TCSCommand.track) OR
	(bGoHomeActive AND eExcludeOwn <> E_TCSCommand.gohome) OR
	TCS_command = E_TCSCommand.goto OR TCS_command = E_TCSCommand.slew OR TCS_command = E_TCSCommand.track OR
	bTracking OR bMoveAbortPending;
END_METHOD

// TRUE if the move may run (accepted, or it replaces the running one), FALSE if it was rejected (logged by the body, nothing written).
// A replace asks for the supersede block of the body: the others are dropped, the axes stopped, the kept move starts at standstill.
METHOD PROTECTED _AcceptMove : BOOL
VAR_INPUT
	eCommand	: E_TCSCommand;
	eExcludeOwn	: E_TCSCommand;
END_VAR
VAR
	eReason		: BROTLib.E_CommandRejectReason;
	eDecision	: BROTLib.E_CommandDecision;
END_VAR
eDecision := BROTLib.F_CommandAcceptance(eCommand := eCommand, stState := _CommandState(eExcludeOwn := eExcludeOwn), eReason => eReason);
IF eDecision = BROTLib.E_CommandDecision.reject THEN
	_NoteRejected(eCommand := eCommand, eReason := eReason);
	_AcceptMove := FALSE;
ELSE
	IF eDecision = BROTLib.E_CommandDecision.replace THEN
		bSupersedeRequest := TRUE;
		eSupersedeKeep := eCommand;
	END_IF
	_AcceptMove := TRUE;
END_IF
END_METHOD

METHOD PRIVATE _NoteRejected
VAR_INPUT
	eCommand	: E_TCSCommand;
	eReason		: BROTLib.E_CommandRejectReason;
END_VAR
nCommandRejectCount := nCommandRejectCount + 1;
eLastRejectedCommand := eCommand;
eLastRejectReason := eReason;
bCommandRejected := TRUE;
END_METHOD

// Every automatic stop (horizon, pole zone, no valid time, lost calibration, bad target): a stop, and a park that is only pending
// (not dispatched yet) is queued behind it instead of being cleared by the stop: it runs when the stop has settled (IAG#84).
METHOD PROTECTED _AutoStop
bStopActive := TRUE;
IF bParkActive AND TCS_command <> E_TCSCommand.park THEN
	bParkAfterStop := TRUE;
	bParkActive := FALSE;
END_IF
END_METHOD

// The park with an error, an E-stop or the axes off: what is safe without the mount (covers, dome, focus), moved unchanged out of the
// arbitration chain (command model step 3C.2). Clears bParkActive, sets bSafeParked for an axes-off park, TCS_command no_command.
METHOD PRIVATE _ParkInPlace
		// Park during an error: the axes are disabled by the error and the park state machine aborts on bError, so
		// bPark used to stay set and the park fired after the next Init() (or hung half way after a reset). Do what
		// is safe without the mount: close the covers, park the dome, disable the focus, and drop the command. The
		// mount is not moved and bIsParked is not set.
		// The same with the axes off (#54): the park command is dispatched only with bReady, which needs the axes
		// enabled, so a park after a stopped power-on, or on a parked telescope, waited until a power-on or the
		// 600 s timeout with the covers open. Not while a park is running (TCS_command park): stage 60 of the park
		// disables the axes itself and the park must go on to stage 100.
		// An E-stop (#57) aborts a running park at any stage: after stage 60 the axes are off and no NC error is raised,
		// so bError stayed FALSE and the park waited at stage 90 for covers that cannot move, until the 600 s timeout.
		bGoHomeActive := FALSE;
		sHomeEnd := 'cancelled by park';
		bGotoActive := FALSE;
		bSlewActive := FALSE;
		bInterrupted := TRUE;
		_ParkTelescope();
		_HomeTelescope();
		_GotoTelescope();
		_SlewTelescope();
		bInterrupted := FALSE;
		fbCovers.Close();
		fbDome.Position := 180.0;
		fbDome.Park();
		IF fbFocus <> 0 THEN
			fbFocus.Enable := FALSE;
		END_IF
		bParkActive := FALSE;
		// #57: say what was commanded, not what was done. With the E-stop pressed the cover and dome requests are
		// dropped; a dome in its latched error ignores the park.
		IF bEstopTriggered THEN
			sParkWhy := 'E-stop pressed, the covers and the dome cannot move. Release it, reset, then park again.';
		ELSE
			IF fbCovers.Closed THEN
				sParkWhy := 'covers closed, ';
			ELSE
				sParkWhy := 'covers closing, ';
			END_IF
			IF fbDome.Error THEN
				sParkWhy := CONCAT(sParkWhy, 'the dome is in error and not parked, ');
			ELSE
				sParkWhy := CONCAT(sParkWhy, 'dome parking, ');
			END_IF
			IF bParkLogged THEN
				sParkWhy := CONCAT(sParkWhy, 'the mount stopped short of the park position');
			ELSE
				sParkWhy := CONCAT(sParkWhy, 'the mount was not moved');
			END_IF
			IF bError THEN
				sParkWhy := CONCAT(sParkWhy, '. Reset, then park again.');
			ELSE
				sParkWhy := CONCAT(sParkWhy, '.');
			END_IF
		END_IF
		IF bParkLogged THEN
			// A running park ends with ONE line, the PARK line, at WARN (E8 logged "PARK completed" and "Park refused").
			IF bEstopTriggered THEN
				sParkEnd := CONCAT('aborted: ', sParkWhy);
				TCSparkEvent.OffLevel := ADSLOG_MSGTYPE_WARN;
			ELSIF bError THEN
				sParkEnd := CONCAT('aborted by an error: ', sParkWhy);
				TCSparkEvent.OffLevel := ADSLOG_MSGTYPE_WARN;
			ELSE
				// #197/#200: the park goes on as an in-place park (covers, dome); its end is this park's one end line
				bParkInPlaceOpen := TRUE;
			END_IF
		ELSE
			// A request during an error or with the axes off was never logged: the separate WARN.
			IF bEstopTriggered THEN
				TCSparkErrorEvent.OnMessage := CONCAT('Park refused: ', sParkWhy);
			ELSIF bError THEN
				TCSparkErrorEvent.OnMessage := CONCAT('Park during an error: ', sParkWhy);
			ELSE
				TCSparkErrorEvent.OnMessage := CONCAT('Park with the axes off: ', sParkWhy);
			END_IF
			bParkInError := TRUE;
		END_IF
		// #110/#187: with no error and no E-stop this leaves a known, covered state. READY_STATE reports 0.3 while the covers
		// close, and bIsParked is set once the covers are closed and the dome is parked (see below); the mount is where it was.
		bSafeParked := NOT bError AND NOT bEstopTriggered;
		TCS_command := E_TCSCommand.no_command;
END_METHOD

// plan step 3.4: the reset trigger and the reset handling of the body (bResetActive, drop of pending goto/slew/track, dome reset, stage reset), moved
// unchanged; called where the block stood. The axis reset of #11 stays in the body, it runs after the error ID.
METHOD PROTECTED _HandleReset
VAR_INPUT
END_VAR
// set reset state either by hardware (key pressed) or by software (set by e.g. tcs)
// #36: the request from Reset() must not be overwritten by the key state, so it has its own flag
// #59: also while the safety acknowledge after an E-stop is pending, so a reset sent during the E-stop (which
// clears the axis errors but skips the acknowledge) or after an E-stop without an axis error is not lost
rtrigResetAny(CLK := fbCabinet.Reset OR bResetRequest);
rtrigReset(CLK := (fbCabinet.Reset OR bResetRequest) AND (bError OR bSafetyAckPending), Q=>bResetActive);
bResetRequest := FALSE;

// The request part of the reset runs on every reset edge, also without an error (MONETcommon#84/#85): pending moves are dropped,
// a move that is still running is stopped (abort stop), a power-on that is running is aborted. The hardware part below (safety
// acknowledge, axis reset passes, dome reset, coordinates) stays gated on an error or a pending acknowledge (#36, #59).
IF rtrigResetAny.Q THEN
	bSupersedeRequest := FALSE;
	bGotoActive := FALSE;
	bSlewActive := FALSE;
	bTrackActive := FALSE;
	bInterrupted := TRUE;
	_GotoTelescope();
	_SlewTelescope();
	IF NOT bLimitHome THEN	// the home of a park in a limit belongs to the park (#84)
		bGoHomeActive := FALSE;
		sHomeEnd := 'cancelled by reset';
		_HomeTelescope();
	END_IF
	bInterrupted := FALSE;
	// a stop that is stuck in Stopping is recovered by a reset without writing over ADS: only axes that stand still are reset (a reset
	// under motion was followed by 0x4260, MONETcommon#84), a moving enabled axis keeps the stop going (MONETcommon#96 D3)
	IF (bStopActive OR bMoveAbortPending)
		AND NOT (fbHourAngle.bEnable AND (aAxis[1].bInMotion OR aAxis[1].bInRamp))
		AND NOT (fbDeclination.bEnable AND (aAxis[2].bInMotion OR aAxis[2].bInRamp)) THEN
		IF aAxis[1].bStopping THEN
			fbHourAngle.Reset();
		END_IF
		IF aAxis[2].bStopping THEN
			fbDeclination.Reset();
		END_IF
		fbStopTx.Cancel();	// the stop then releases at standstill
	END_IF
	// not during an error (the drives are off) and not during a park (its motion is wanted)
	bMoveAbortPending := bMoveAbortPending OR BROTLib.F_ResetMoveAbort(
		bError := bError,
		bParkRunning := TCS_command = E_TCSCommand.park,
		bAnyAxisMoving := (fbHourAngle.bEnable AND (aAxis[1].bInMotion OR aAxis[1].bInRamp OR aAxis[1].bHoming))
			OR (fbDeclination.bEnable AND (aAxis[2].bInMotion OR aAxis[2].bInRamp OR aAxis[2].bHoming)));
	IF bPowerActive OR fbStartup.Initializing THEN
		bStopActive := TRUE;	// aborts the power-on and marks the startup aborted (stop branch)
	END_IF
END_IF

IF bResetActive THEN
    fbStartup.MarkAborted();
	bTestError := FALSE;
	bSoftwareError := FALSE;
	nSoftwareErrorID := 0;
	// reset input coords to parking position (always over horizon to stop bHorizonError from occuring)
	fDeclination := telescopeConfig.declinationPark;
	fbHaDec2RaDec(	jd := fJd +fTimeOffset,
					ha := telescopeConfig.houranglePark,
					dec := telescopeConfig.declinationPark,
					lon := telescopeConfig.longitude,
					ra_out => fRightAscension);
	// reset elevation values to abitrarry value over horizon, will get overwritten down the line
	fElevationCalc := 20.0;
	fElevation := 20.0;
	// reset dome position
	fbDome.Position := 180.0;
	// #35: a dome error after an E-stop (serial link lost) stays latched until the dome is reset, and nothing else
	// reaches it. Only the dome's error state reacts to a reset; in every other state it is ignored.
	IF fbDome <> 0 THEN
		fbDome.Reset();
	END_IF
	// reset the stages of all statemachine methods
	// #100: a goto/slew/track request that is still pending must not outlive the reset (the error clears them only
	// while it lasts)
	bGotoActive := FALSE;
	bSlewActive := FALSE;
	bTrackActive := FALSE;
	bInterrupted := TRUE;
	_HomeTelescope();
	_GotoTelescope();
	_SlewTelescope();
	_ParkTelescope();
	bInterrupted := FALSE;
END_IF
END_METHOD

// plan step 3.2: the feedback of the two axes (the outputs of their FB_Axis) once per scan, at the start of the body. The outputs
// do not change while the telescope body runs, so they are the same wherever the body reads them.
METHOD PRIVATE _ReadAxes
VAR_INPUT
END_VAR
aAxis[1].bStandStill := fbHourAngle.fbAxis.StandStill;
aAxis[1].bStopDone := fbHourAngle.fbAxis.StopDone;
aAxis[1].bInMotion := fbHourAngle.fbAxis.InMotion;
aAxis[1].bInRamp := fbHourAngle.fbAxis.InRamp;
aAxis[1].bHoming := fbHourAngle.fbAxis.Homing;
aAxis[1].bStopping := fbHourAngle.fbAxis.Stopping;
aAxis[1].bBusy := fbHourAngle.fbAxis.Busy;
aAxis[1].bTracking := fbHourAngle.fbAxis.isTracking;
aAxis[2].bStandStill := fbDeclination.fbAxis.StandStill;
aAxis[2].bStopDone := fbDeclination.fbAxis.StopDone;
aAxis[2].bInMotion := fbDeclination.fbAxis.InMotion;
aAxis[2].bInRamp := fbDeclination.fbAxis.InRamp;
aAxis[2].bHoming := fbDeclination.fbAxis.Homing;
aAxis[2].bStopping := fbDeclination.fbAxis.Stopping;
aAxis[2].bBusy := fbDeclination.fbAxis.Busy;
aAxis[2].bTracking := fbDeclination.fbAxis.isTracking;
END_METHOD

METHOD PRIVATE _GotoTelescope : USINT
VAR_INPUT
END_VAR
VAR
	GoToEvent		: FB_Eventlog;
END_VAR
VAR_INST
	nStage			: USINT := 0;
	nLastStage		: USINT := 101;
END_VAR
_GotoTelescope := nStage;
IF tonGotoTimeout.Q THEN	// MONETcommon#17: fed every scan in the body, a method-local TON never kept its state
	bSoftwareError := TRUE;		// #30: latched until a reset, bError is recomputed every scan
	nSoftwareErrorID := 16#10;
	bGotoActive := FALSE;
	nStage := 0;
	RETURN;
END_IF
IF bResetActive OR bError OR bStopActive OR bInterrupted THEN
	nStage := 0;
	RETURN;
END_IF

CASE nStage OF
	0:	
		IF bReady AND NOT bBusy THEN
			nStage := 10;
		END_IF
	10:
		IF fbHourAngle.Tracking = TRUE OR fbDeclination.Tracking = TRUE THEN
			fbHourAngle.Tracking := FALSE;
			fbDeclination.Tracking := FALSE;
		ELSE
			nStage := 20;
		END_IF
	20:
		// send Dome position
		THIS^.fbDome.Position := fAzimuthCalc;
		// clear offsets
		THIS^.HourAngleOffset := 0.0;
		THIS^.DeclinationOffset := 0.0;
		// Declination (including offest and pointing model)
		fbDeclination.Position := fDeclinationApparent + fDeclinationOffset + fDeclinationPointingOffset;
		// HourAngle
		// change to -180 to 180 degree in HA
		IF MODABS(fHourAngleApparent + F_HourAngleOffsetOnAxis(fHourAngleOffset, fDeclinationApparent)+ fHourAnglePointingOffset, 360) > 180 THEN
			fbHourAngle.Position := MODABS(fHourAngleApparent + F_HourAngleOffsetOnAxis(fHourAngleOffset, fDeclination)+ fHourAnglePointingOffset,360) - 360.0;
		ELSE
			fbHourAngle.Position := MODABS(fHourAngleApparent + F_HourAngleOffsetOnAxis(fHourAngleOffset, fDeclination)+ fHourAnglePointingOffset,360);
		END_IF


		fbHourAngle.Velocity := fSlewVelocity;
		fbDeclination.Velocity := fSlewVelocity;
		
		// make sure to never drive under Horizon
		IF ABS(fbHourAngle.Position) < ABS(fHourAngleCurrent) THEN
			// move Ha then Dec
			nStage := 30;
		ELSE
			// move Dec then HA
			nStage := 40;
		END_IF
	// Stage 30: move Ha and then Dec
	30:
		fbHourAngle.MoveAxis := TRUE;
		IF fbHourAngle.Busy THEN
			nStage := 31;
		END_IF
	31:
		IF NOT fbHourAngle.Busy AND fbHourAngle.MoveDone THEN
			fbHourAngle.MoveAxis := FALSE;
		END_IF
		IF NOT fbHourAngle.MoveAxis THEN
		   nStage := 32;
		END_IF
	32:
		fbDeclination.MoveAxis := TRUE;
		IF fbDeclination.Busy THEN
			nStage := 33;
		END_IF
	33:
		IF NOT fbDeclination.Busy AND fbDeclination.MoveDone THEN
			fbDeclination.MoveAxis := FALSE;
		END_IF
		IF NOT fbDeclination.MoveAxis THEN
		   nStage := 75;
		END_IF
	// Stage 40: move Dec and then Ha
	40:
		fbDeclination.MoveAxis := TRUE;
		IF fbDeclination.Busy THEN
			nStage := 41;
		END_IF
	41:
		IF NOT fbDeclination.Busy AND fbDeclination.MoveDone THEN
			fbDeclination.MoveAxis := FALSE;
		END_IF
		IF NOT fbDeclination.MoveAxis THEN
		   nStage := 42;
		END_IF
	42:
		fbHourAngle.MoveAxis := TRUE;
		IF fbHourAngle.Busy THEN
			nStage := 43;
		END_IF
	43:
		IF NOT fbHourAngle.Busy AND fbHourAngle.MoveDone THEN
			fbHourAngle.MoveAxis := FALSE;
		END_IF
		IF NOT fbHourAngle.MoveAxis THEN
		   nStage := 75;
		END_IF

	75:
		IF NOT bSliding AND bStopped THEN // all axis standstill
			nStage := 100;
		END_IF
	100:
		bGotoActive := FALSE;
		// enable automatic tracking
		bTrackActive := bAutoTrack;
		nStage := 0;
END_CASE
GoToEvent(Trigger := nStage > nLastStage, FormatString := 'GOTO progress: %s', OnMessage := USINT_TO_STRING(nStage), comm := fbComm);
nLastStage := nStage;
END_METHOD

METHOD PRIVATE _HomeTelescope : USINT
VAR_INPUT
END_VAR
VAR
	HomeEvent:	FB_Eventlog;
END_VAR
VAR_INST
	nStage:		USINT := 0;
	nLastStage:	USINT := 101;
END_VAR
_HomeTelescope := nStage;
IF tonHomeTimeout.Q THEN
    fbStartup.MarkAbortedIfInitializing();	// MONETcommon#17: fed every scan in the body
	bSoftwareError := TRUE;		// #30
	nSoftwareErrorID := 16#30;
	bGoHomeActive := FALSE;	// like goto/slew; otherwise the expired timer would fire again right away
	sHomeEnd := 'timed out';
	nStage := 0;
	RETURN;		// #75: like goto/slew/park; bError is recomputed next scan, do not run the stages on
END_IF

IF bResetActive OR bError OR bStopActive OR bInterrupted THEN
    fbStartup.MarkAbortedIfInitializing();
	nStage := 0;
	RETURN;
END_IF
CASE nStage OF
	0:	
		IF bReady AND bSettled AND NOT bBusy THEN
			nStage := 10;
		END_IF
	10:
		IF fbHourAngle.Tracking = TRUE OR fbDeclination.Tracking = TRUE THEN
			fbHourAngle.Tracking := FALSE;
			fbDeclination.Tracking := FALSE;
		ELSE
			nStage := 20;
		END_IF
	20:
		fbHourAngle.Position := telescopeConfig.hourangleHome;
		fbHourAngle.Velocity := fSlewVelocity;
		fbDeclination.Position := telescopeConfig.declinationHome;
		fbDeclination.Velocity := fSlewVelocity;
		
		// make sure to never drive under Horizon
		IF ABS(telescopeConfig.hourangleHome) < ABS(fHourAngleCurrent) THEN
			// move Ha then Dec
			nStage := 30;
		ELSE
			// move Dec then HA
			nStage := 40;
		END_IF
	// nStage 30: move Ha and then Dec
	30:
		fbHourAngle.MoveAxis := TRUE;
        nStage := 31;
	31:
		IF NOT fbHourAngle.Busy AND fbHourAngle.MoveDone THEN
			fbHourAngle.MoveAxis := FALSE;
		END_IF
		IF NOT fbHourAngle.MoveAxis THEN
		   nStage := 32;
		END_IF
	32:
		fbDeclination.MoveAxis := TRUE;
        nStage := 33;
	33:
		IF NOT fbDeclination.Busy AND fbDeclination.MoveDone THEN
			fbDeclination.MoveAxis := FALSE;
		END_IF
		IF NOT fbDeclination.MoveAxis THEN
		   nStage := 100;
		END_IF
	// nStage 40: move Dec and then Ha
	40:
		fbDeclination.MoveAxis := TRUE;
        nStage := 41;
	41:
		IF NOT fbDeclination.Busy AND fbDeclination.MoveDone THEN
			fbDeclination.MoveAxis := FALSE;
		END_IF
		IF NOT fbDeclination.MoveAxis THEN
		   nStage := 42;
		END_IF
	42:
		fbHourAngle.MoveAxis := TRUE;
        nStage := 43;
	43:
		IF NOT fbHourAngle.Busy AND fbHourAngle.MoveDone THEN
			fbHourAngle.MoveAxis := FALSE;
		END_IF
		IF NOT fbHourAngle.MoveAxis THEN
		   nStage := 100;
		END_IF
	100:
        IF fbFocus <> 0 THEN
            fbFocus.Position := telescopeConfig.focusHome;
        END_IF
        IF fbStartup.Initializing AND NOT bParkAfterHome THEN	// #84: a park follows, the startup was aborted
            // Only initialization waits for its remaining focus work; manual Home semantics stay unchanged.
            nStage := 110;
        ELSE
            fRightAscension := fRightAscensionCurrentICRS;
            fDeclination := fDeclinationCurrentICRS;
            bParkHomeDone := bParkAfterHome;	// #84
            bGoHomeActive := FALSE;
            nStage := 0;
        END_IF
    110:
        // Compare with the effective target (the focus applies configured limits). Busy alone has an idle gap
        // between assigning a target and the focus block starting its move. No sampled moving edge is required.
        IF (fbFocus <> 0 AND_THEN (fbFocus.Calibrated AND fbFocus.Ready AND NOT fbFocus.Busy AND
            ABS(fbFocus.Position - fbFocus.ActualPosition) <= fStartupFocusTolerance)) AND bReady AND bMainReady AND bStopped AND NOT bBusy THEN
            fRightAscension := fRightAscensionCurrentICRS;
            fDeclination := fDeclinationCurrentICRS;
            fbStartup.MarkCompleted();
            bGoHomeActive := FALSE;
            nStage := 0;
        END_IF
END_CASE

HomeEvent(Trigger := nStage > nLastStage, FormatString := 'GOHOME progress: %s', OnMessage := USINT_TO_STRING(nStage), comm := fbComm);
nLastStage := nStage;
END_METHOD

METHOD PRIVATE _ParkTelescope : USINT
VAR_INPUT
END_VAR
VAR
	ParkEvent	: FB_Eventlog;
	bFocusMoving	: BOOL;
END_VAR
VAR_INST
	nStage		: USINT := 0;
	nLastStage	: USINT := 0;
END_VAR
_ParkTelescope := nStage;
IF tonParkTimeout.Q THEN	// fed every scan in the body, like the goto/home/slew timeouts
	bSoftwareError := TRUE;
	nSoftwareErrorID := 16#20;
	bParkActive := FALSE;
	sParkEnd := 'timed out';
	nStage := 0;
	RETURN;
END_IF
IF bResetActive OR bError OR bStopActive OR bInterrupted THEN
	nStage := 0;
	RETURN;
END_IF
IF bIsParked THEN
	nStage := 100;
END_IF
CASE nStage OF
	0: 
		IF fbFocus <> 0 THEN
			fbFocus.Position := telescopeConfig.focusPark;
		END_IF
		// (the former "emergency park" under IF bError never ran: the method returns on bError above, and the
		// command is not even started while bError; a park during an error is handled in the arbitration)
		IF NOT bBusy THEN
			nStage := 10;
		END_IF
	10:
		fbDome.StopTrack();
		fbDome.Position := 180.0;
		IF fbHourAngle.Tracking = TRUE OR fbDeclination.Tracking = TRUE THEN
			fbHourAngle.Tracking := FALSE;
			fbDeclination.Tracking := FALSE;
		ELSE
			nStage := 20;
		END_IF
	20:
		fbDome.Park();
		THIS^.HourAngleOffset := 0.0;
		THIS^.DeclinationOffset := 0.0;
		fbHourAngle.Position := telescopeConfig.houranglePark;
		fbHourAngle.Velocity := fSlewVelocity;
		fbDeclination.Position := telescopeConfig.declinationPark;
		fbDeclination.Velocity := fSlewVelocity;
		
		// make sure to never drive under Horizon
		IF ABS(telescopeConfig.houranglePark) < ABS(fHourAngleCurrent) THEN
			// move Ha then Dec
			nStage := 30;
		ELSE
			// move Dec then HA
			nStage := 40;
		END_IF
	// Stage 30: move Ha and then Dec
	30:
		fbHourAngle.MoveAxis := TRUE;
		IF fbHourAngle.Busy THEN
			nStage := 31;
		END_IF
	31:
		IF NOT fbHourAngle.Busy AND fbHourAngle.MoveDone THEN
			fbHourAngle.MoveAxis := FALSE;
		END_IF
		IF NOT fbHourAngle.MoveAxis THEN
		   nStage := 32;
		END_IF
	32:
		fbDeclination.MoveAxis := TRUE;
		IF fbDeclination.Busy THEN
			nStage := 33;
		END_IF
	33:
		IF NOT fbDeclination.Busy AND fbDeclination.MoveDone THEN
			fbDeclination.MoveAxis := FALSE;
		END_IF
		IF NOT fbDeclination.MoveAxis THEN
		   nStage := 60;
		END_IF
	// Stage 40: move Dec and then Ha
	40:
		fbDeclination.MoveAxis := TRUE;
		IF fbDeclination.Busy THEN
			nStage := 41;
		END_IF
	41:
		IF NOT fbDeclination.Busy AND fbDeclination.MoveDone THEN
			fbDeclination.MoveAxis := FALSE;
		END_IF
		IF NOT fbDeclination.MoveAxis THEN
		   nStage := 42;
		END_IF
	42:
		fbHourAngle.MoveAxis := TRUE;
		IF fbHourAngle.Busy THEN
			nStage := 43;
		END_IF
	43:
		IF NOT fbHourAngle.Busy AND fbHourAngle.MoveDone THEN
			fbHourAngle.MoveAxis := FALSE;
		END_IF
		IF NOT fbHourAngle.MoveAxis THEN
		   nStage := 60;
		END_IF
	60:
		IF NOT fbHourAngle.Enable AND NOT fbDeclination.Enable THEN
			// #66: request the close once; repeating it every scan latched bClose in FB_CoverControl
			fbCovers.Close();
			nStage := 80;
		END_IF

		IF bStopped THEN
			fbHourAngle.Enable := FALSE;
			fbDeclination.Enable := FALSE;
		END_IF
		
		fbHourAngle.MoveAxis := FALSE;
		fbDeclination.MoveAxis := FALSE;
	80:
		// (the former "IF an axis is enabled THEN nStage := 60" was overwritten by the line below and never took
		// effect; nothing enables an axis while the park runs, _PowerOn is a different command)
		// #56: the focus move to focusPark starts at stage 0. A park from home does not move the mount, so the axes
		// are off after about a second and the focus enable was removed while it was still moving (error 16992
		// "Controller enable"). Wait until it has arrived or stopped (at most 60 s), then disable it.
		bFocusMoving := fbFocus <> 0 AND_THEN (fbFocus.Calibrated AND (fbFocus.Busy OR ABS(fbFocus.Position - fbFocus.ActualPosition) > 0.05));
		tonParkFocus(IN := bFocusMoving, PT := T#60S, nDivisor := nTimeDivisor);
		IF NOT bFocusMoving OR tonParkFocus.Q THEN
			IF fbFocus <> 0 THEN
				fbFocus.Enable := FALSE;
			END_IF
			tonParkFocus(IN := FALSE);
			nStage := 90;
		END_IF
	90:
		IF fbCovers.Closed THEN
			nStage := 100;
		END_IF
	100:
		bIsPowered:=FALSE;
		bIsParked := TRUE;
		bParkedInPlace := FALSE;
		bParkActive := FALSE;
		_ParkTelescope := 100;
		nStage := 0;	
END_CASE
ParkEvent(Trigger := nStage > nLastStage, FormatString := 'Parking progress: %s', OnMessage := USINT_TO_STRING(nStage), comm := fbComm);
nLastStage := nStage;
END_METHOD

// #11: reset every axis that has an error, also a hidden one (nErrorID set with the error flag FALSE)
METHOD PRIVATE _ResetErroredAxes
VAR_INPUT
	bAll	: BOOL;		// also reset axes that are not enabled (#55), the second pass after the acknowledge
END_VAR
IF fbHourAngle.Error OR fbHourAngle.nErrorID <> 0 OR (bAll AND NOT fbHourAngle.Enable) THEN
	fbHourAngle.Reset();
END_IF
IF fbDeclination.Error OR fbDeclination.nErrorID <> 0 OR (bAll AND NOT fbDeclination.Enable) THEN
	fbDeclination.Reset();
END_IF
IF fbFocus <> 0 AND_THEN (fbFocus.Error OR fbFocus.ErrorID <> 0 OR (bAll AND NOT fbFocus.Enable)) THEN
	fbFocus.Reset();
END_IF
END_METHOD

// #39: the reason a power-on cannot start, as one line for the ADS log. First match wins.
METHOD PRIVATE _PowerOnBlockedReason : STRING(120)
VAR
	sAxis		: STRING(8);
	nId			: UDINT;
END_VAR
IF bEstopTriggered THEN
	_PowerOnBlockedReason := 'Power-on blocked: E-stop pressed. Release it, then reset.';
	RETURN;
END_IF

// the axis ids are used even when bError is FALSE (a hidden NC error, HA 16933 on 2026-10-12)
IF fbHourAngle.nErrorID <> 0 THEN
	sAxis := 'HA';
	nId := fbHourAngle.nErrorID;
ELSIF fbDeclination.nErrorID <> 0 THEN
	sAxis := 'Dec';
	nId := fbDeclination.nErrorID;
ELSIF fbFocus <> 0 AND_THEN fbFocus.ErrorID <> 0 THEN
	sAxis := 'Focus';
	nId := fbFocus.ErrorID;
END_IF

IF nId <> 0 THEN
	IF nId = 18000 OR nId = 19209 THEN
		// drive hardware not ready / axis not ready: the drives are in STO until the safety is acknowledged
		_PowerOnBlockedReason := CONCAT(CONCAT(CONCAT(CONCAT('Power-on blocked: safety not acknowledged (', sAxis), ' '), UDINT_TO_STRING(nId)), '). Reset the telescope (cabinet key or reset command).');
	ELSE
		_PowerOnBlockedReason := CONCAT(CONCAT(CONCAT(CONCAT('Power-on blocked: ', sAxis), ' error '), UDINT_TO_STRING(nId)), '. Reset the telescope.');
	END_IF
ELSIF bSafetyAckPending THEN
	_PowerOnBlockedReason := 'Power-on blocked: safety not acknowledged after the E-stop. Reset the telescope (cabinet key or reset command).';
ELSIF bSoftwareError THEN
	_PowerOnBlockedReason := CONCAT(CONCAT('Power-on blocked: command timeout error ', UDINT_TO_STRING(nSoftwareErrorID)), '. Reset the telescope.');
ELSE
	_PowerOnBlockedReason := 'Power-on blocked: telescope error. Reset the telescope.';
END_IF
END_METHOD

METHOD PRIVATE _PowerOn : USINT
VAR_INPUT
END_VAR
VAR
	PowerOnEvent	: FB_Eventlog;
END_VAR
VAR_INST
	nStage		: USINT := 0;
	nLastStage	: USINT := 0;
	tonCalibTimeout	: TON;		// #155: stage 40 had no timeout
END_VAR
// #59: also refused while the safety acknowledge after an E-stop is pending. While the reset is running
// (bAxisResetAfterAck) the power-on waits at stage 0 as before; the acknowledge ends before that wait does.
IF bError OR (bSafetyAckPending AND NOT bAxisResetAfterAck) THEN
	bPowerFailure := TRUE;
	TCSpowerEvent.OnMessage := 'failed';
	// #39: say why, on every refused request. bPowerFailure stays TRUE until a power-on succeeds, so it gives
	// no new edge for the second request and logged nothing; this one-scan flag does.
	TCSpowerBlockedEvent.OnMessage := _PowerOnBlockedReason();
	bPowerBlocked := TRUE;
	bPowerActive := FALSE;
ELSE
	bPowerFailure := FALSE;		
END_IF

_PowerOn := nStage;
// #69: a power-on only runs while it is requested. Stage 100 clears bPower, but TCS_command stays poweron until
// the go-home takes over, so _PowerOn kept being called and restarted its stages; the go-home then left nStage at
// 10 or 20 and the next power=1 resumed there, skipping the wait for the safety acknowledge in stage 0.
IF NOT bPowerActive OR bResetActive OR bError OR bStopActive OR bInterrupted THEN
    // After a successful handoff bPower is false but the home phase still owns startup.
    IF bResetActive OR bError OR bStopActive OR bInterrupted OR bPowerFailure THEN
        fbStartup.MarkAborted();
        bPowerActive := FALSE;
    END_IF
	nStage := 0;
	nLastStage := 0;	// #195: else the stages up to the aborted one are not logged in the next power-on
	RETURN;
END_IF

IF nStage >= 40 THEN
    fbStartup.MarkCalibrating();
END_IF

// #155: an axis that never starts its calibration (no error, no log) held the power-on in stage 40 for good. The sweep
// of one axis takes about 35 s; end the power-on as a failed startup if it lasts three minutes.
tonCalibTimeout(IN := nStage = 40, PT := T#3M);
IF tonCalibTimeout.Q THEN
	bPowerFailure := TRUE;
	TCSpowerEvent.OnMessage := 'failed';
	IF fbHourAngle.Calibrated THEN
		TCSpowerBlockedEvent.OnMessage := 'POWER: calibration timeout (Declination is not calibrated)';
	ELSIF fbDeclination.Calibrated THEN
		TCSpowerBlockedEvent.OnMessage := 'POWER: calibration timeout (Hour Angle is not calibrated)';
	ELSE
		TCSpowerBlockedEvent.OnMessage := 'POWER: calibration timeout (neither axis is calibrated)';
	END_IF
	bPowerBlocked := TRUE;
	fbStartup.MarkAborted();
	bPowerActive := FALSE;
	nStage := 0;
	nLastStage := 0;	// #195
	RETURN;
END_IF

CASE nStage OF
	0:
		// #55: wait for the axis reset that follows the safety acknowledge (at most 2.5 s); enabling the axes before
		// it gave 18000 on HA and Dec
		IF NOT bAxisResetAfterAck THEN
			bIsParked := FALSE;
			bParkedInPlace := FALSE;
			IF bCoverAutoOpen THEN
				// check if covers should automatic open
				nStage := 10;
			ELSE
				nStage := 40;
			END_IF
		END_IF
	10:
		// COVER MUST BE OPENED FOR A SUCCESSFUL WAKE & SHAKE COMMAND!
		IF NOT fbCovers.Opened THEN
			fbCovers.Open();
		END_IF
		nStage := 20;
	20:
		IF bMainReady AND fbCovers.Opened THEN
			nStage := 40;
		END_IF
	40:
		// enable hourangle, enable declination
		// #69: never while the safety acknowledge runs (the drives are still in STO: 0x441C, then 4225 on HA)
		IF NOT bAxisResetAfterAck THEN
			fbHourAngle.Enable := TRUE;
			fbDeclination.Enable := TRUE;
			// #100/#103: calibration alone is not enough. The NC keeps Homed through a Reset Cold while the drives are
			// still in STO, so stages 40, 70 and 100 ran in consecutive scans before the enable failed (18000): stage 100
			// set bIsPowered and the go-home, bReady pulsed ("startup finished") and the error left bIsPowered TRUE.
			// Wait for the power status of both axes (MC_Power Status); an enable error ends the power-on above.
			IF fbHourAngle.bReady AND fbDeclination.bReady AND fbHourAngle.Calibrated AND fbDeclination.Calibrated THEN
				nStage := 70;
			END_IF
		END_IF
	70:
		// if Focus, enable and calibrate
		IF fbFocus <> 0 THEN
			fbFocus.Enable := TRUE;
			fbFocus.Position := telescopeConfig.focusPark;
			IF fbFocus.Calibrated THEN
				nStage := 100;
			END_IF
		ELSE
			nStage := 100;
		END_IF
	100:
		//PowerOn is done, set bPower to False
		bPowerActive := FALSE;
		bIsPowered := TRUE;
		// slew the telescope to the home position
		bGoHomeActive := TRUE;
		// set dome to tracking
		fbDome.Position := 180.0;// reset Dome position
		fbDome.Track();
		_PowerOn := 100;
		nStage := 0;	
END_CASE
PowerOnEvent(Trigger := nStage > nLastStage, FormatString := 'PowerOn progress: %s', OnMessage := USINT_TO_STRING(nStage), comm := fbComm);
nLastStage := nStage;
END_METHOD

METHOD _SendTelemetryEquitorial : BOOL
VAR_INPUT

END_VAR
(* Open TSI / TCI standart *)

(* TELESCOPE module*)

fbComm.PublishLREAL('telescope', 'dome', 'TELESCOPE.READY_STATE',	fReadyState);
fbComm.PublishLREAL('telescope', 'dome', 'TELESCOPE.MOTION_STATE',	nMotionState);

// INFO
fbComm.PublishString('telescope', 'dome', 'TELESCOPE.INFO.NAME',	telescopeConfig.name);
fbComm.PublishLREAL('telescope', 'dome', 'TELESCOPE.INFO.DIAMETER',	telescopeConfig.diameter);
fbComm.PublishString('telescope', 'dome', 'TELESCOPE.INFO.CABINET',	telescopeConfig.cabinet);
fbComm.PublishString('telescope', 'dome', 'TELESCOPE.INFO.MANUFACTURER', telescopeConfig.manufacturer);

// CONFIG
IF fbDome <> 0 THEN
	fbComm.PublishINT('telescope', 'dome', 'TELESCOPE.CONFIG.CAPABILITIES', fbDome.Capabilities);
ELSE
	fbComm.PublishINT('telescope', 'dome', 'TELESCOPE.CONFIG.CAPABILITIES', 0);
END_IF
fbComm.PublishString('telescope', 'dome', 'TELESCOPE.CONFIG.MOUNTOPTIONS', telescopeConfig.mountOptions);
fbComm.PublishString('telescope', 'dome', 'TELESCOPE.CONFIG.MOUNT', telescopeConfig.mount);

// STATUS
IF bEstopTriggered THEN
	fbComm.PublishINT('telescope', 'dome', 'TELESCOPE.STATUS.GLOBAL', 1);
ELSIF bError THEN
	fbComm.PublishINT('telescope', 'dome', 'TELESCOPE.STATUS.GLOBAL', 2);
ELSE
	fbComm.PublishINT('telescope', 'dome', 'TELESCOPE.STATUS.GLOBAL', 0);
END_IF

IF bLocalMode THEN
	fbComm.PublishINT('telescope', 'dome', 'TELESCOPE.STATUS.LOCAL_MODE', 1);
ELSE
	fbComm.PublishINT('telescope', 'dome', 'TELESCOPE.STATUS.LOCAL_MODE', 0);
END_IF
(* ERROR LIST: TO BE IMPLEMENTED!!!*)

(* OBJECT Module*)
// Set Coords from outside | GoTo:RA DEC | Slew:Alt Az

// INSTRUMENTAL
fbComm.PublishLREAL('telescope', 'dome', 'OBJECT.INSTRUMENTAL.DEC', fDeclinationApparent + fDeclinationOffset + fDeclinationPointingOffset);
// change to -180 to 180 degree in HA
IF MODABS(fHourAngleApparent + F_HourAngleOffsetOnAxis(fHourAngleOffset, fDeclination)+ fHourAnglePointingOffset, 360) > 180 THEN
	fbComm.PublishLREAL('telescope', 'dome', 'OBJECT.INSTRUMENTAL.HA', MODABS(fHourAngleApparent + F_HourAngleOffsetOnAxis(fHourAngleOffset, fDeclinationApparent)+ fHourAnglePointingOffset,360)- 360.0);
ELSE
	fbComm.PublishLREAL('telescope', 'dome', 'OBJECT.INSTRUMENTAL.HA', MODABS(fHourAngleApparent + F_HourAngleOffsetOnAxis(fHourAngleOffset, fDeclinationApparent)+ fHourAnglePointingOffset,360));
END_IF

// HORIZONTAL
IF bSlewActive THEN
	fbComm.PublishLREAL('telescope', 'dome', 'OBJECT.HORIZONTAL.ALT', fElevation);
	fbComm.PublishLREAL('telescope', 'dome', 'OBJECT.HORIZONTAL.AZ', fAzimuth);
ELSE
	fbComm.PublishLREAL('telescope', 'dome', 'OBJECT.HORIZONTAL.ALT', fElevationCalc);
	fbComm.PublishLREAL('telescope', 'dome', 'OBJECT.HORIZONTAL.AZ', fAzimuthCalc);
END_IF

//EQUATORIAL
fbComm.PublishString('telescope', 'dome', 'OBJECT.EQUATORIAL.EPOCH', 'J2000.0');
fbComm.PublishString('telescope', 'dome', 'OBJECT.EQUATORIAL.EQUINOX', 'J2000.0');
fbComm.PublishLREAL('telescope', 'dome', 'OBJECT.EQUATORIAL.RA_PM', 0.0);
fbComm.PublishLREAL('telescope', 'dome', 'OBJECT.EQUATORIAL.DEC_PM', 0.0);
fbComm.PublishLREAL('telescope', 'dome', 'OBJECT.EQUATORIAL.RA_RATE', 0.0);
fbComm.PublishLREAL('telescope', 'dome', 'OBJECT.EQUATORIAL.DEC_RATE', 0.0);
fbComm.PublishLREAL('telescope', 'dome', 'OBJECT.EQUATORIAL.RA', fRightAscension);	// degrees (BROTLib#37)
fbComm.PublishLREAL('telescope', 'dome', 'OBJECT.EQUATORIAL.DEC', fDeclination);
fbComm.PublishLREAL('telescope', 'dome', 'OBJECT.EQUATORIAL.HA_APPARENT', fHourAngleApparent);
fbComm.PublishLREAL('telescope', 'dome', 'OBJECT.EQUATORIAL.DEC_APPARENT', fDeclinationApparent);


(* POINTING *)
fbComm.PublishLREAL('telescope', 'dome', 'POINTING.SLEWTIME', fSlewtime);
fbComm.PublishLREAL('telescope', 'dome', 'POINTING.OFFSETS.HA', fHourAnglePointingOffset);
fbComm.PublishLREAL('telescope', 'dome', 'POINTING.OFFSETS.DEC', fDeclinationPointingOffset);


(*POSITION*)
//LOCAL
fbComm.PublishLREAL('telescope', 'dome', 'POSITION.LOCAL.SIDEREAL_TIME', fLst);
fbComm.PublishLREAL('telescope', 'dome', 'POSITION.LOCAL.JD', fJd);
fbComm.PublishLREAL('telescope', 'dome', 'POSITION.LOCAL.LATITUDE', telescopeConfig.latitude);
fbComm.PublishLREAL('telescope', 'dome', 'POSITION.LOCAL.LONGITUDE', telescopeConfig.longitude);
fbComm.PublishLREAL('telescope', 'dome', 'POSITION.LOCAL.HEIGHT', telescopeConfig.altitude);
//INSTRUMENTAL
// > DEC
// POWER_STATE
IF fbDeclination.Enable THEN
	fbComm.PublishLREAL('telescope', 'dome', 'POSITION.INSTRUMENTAL.DEC.POWER_STATE', 1.0);
ELSE
	fbComm.PublishLREAL('telescope', 'dome', 'POSITION.INSTRUMENTAL.DEC.POWER_STATE', 0.0);
END_IF
//REFERENCED
IF fbDeclination.Calibrated THEN
	fbComm.PublishLREAL('telescope', 'dome', 'POSITION.INSTRUMENTAL.DEC.REFERENCED', 1.0);
ELSE
	fbComm.PublishLREAL('telescope', 'dome', 'POSITION.INSTRUMENTAL.DEC.REFERENCED', 0.0);
END_IF
//ERROR_STATE
IF fbDeclination.Error THEN
	fbComm.PublishINT('telescope', 'dome', 'POSITION.INSTRUMENTAL.DEC.ERROR_STATE', fbDeclination.ErrorID);
ELSE
	fbComm.PublishINT('telescope', 'dome', 'POSITION.INSTRUMENTAL.DEC.ERROR_STATE', 0);
END_IF
//MOTION_STATE
IF fbDeclination.Busy THEN
	IF fbDeclination.isTracking THEN
		fbComm.PublishINT('telescope', 'dome', 'POSITION.INSTRUMENTAL.DEC.MOTION_STATE', 8);
	ELSE
		fbComm.PublishINT('telescope', 'dome', 'POSITION.INSTRUMENTAL.DEC.MOTION_STATE', 1);
	END_IF
ELSE
	fbComm.PublishINT('telescope', 'dome', 'POSITION.INSTRUMENTAL.DEC.MOTION_STATE', 0);
END_IF
fbComm.PublishLREAL('telescope', 'dome', 'POSITION.INSTRUMENTAL.DEC.REALPOS', fDeclinationCurrent-fDeclinationOffset);
fbComm.PublishLREAL('telescope', 'dome', 'POSITION.INSTRUMENTAL.DEC.CURRPOS', fDeclinationCurrent);
fbComm.PublishLREAL('telescope', 'dome', 'POSITION.INSTRUMENTAL.DEC.TARGETPOS', fbDeclination.Position);
fbComm.PublishLREAL('telescope', 'dome', 'POSITION.INSTRUMENTAL.DEC.CURRSPEED', fbDeclination.Velocity);
fbComm.PublishLREAL('telescope', 'dome', 'POSITION.INSTRUMENTAL.DEC.TARGETDISTANCE', ABS(fDeclinationCurrent-fbDeclination.Position));
fbComm.PublishLREAL('telescope', 'dome', 'POSITION.INSTRUMENTAL.DEC.OFFSET', fDeclinationOffset);

// > HA
// POWER_STATE
IF fbHourAngle.Enable THEN
	fbComm.PublishLREAL('telescope', 'dome', 'POSITION.INSTRUMENTAL.HA.POWER_STATE', 1.0);
ELSE
	fbComm.PublishLREAL('telescope', 'dome', 'POSITION.INSTRUMENTAL.HA.POWER_STATE', 0.0);
END_IF
//REFERENCED
IF fbHourAngle.Calibrated THEN
	fbComm.PublishLREAL('telescope', 'dome', 'POSITION.INSTRUMENTAL.HA.REFERENCED', 1.0);
ELSE
	fbComm.PublishLREAL('telescope', 'dome', 'POSITION.INSTRUMENTAL.HA.REFERENCED', 0.0);
END_IF
//ERROR_STATE
IF fbHourAngle.Error THEN
	fbComm.PublishINT('telescope', 'dome', 'POSITION.INSTRUMENTAL.HA.ERROR_STATE', fbHourAngle.ErrorID);
ELSE
	fbComm.PublishINT('telescope', 'dome', 'POSITION.INSTRUMENTAL.HA.ERROR_STATE', 0);
END_IF
//MOTION_STATE
IF fbHourAngle.Busy THEN
	IF fbHourAngle.isTracking THEN
		fbComm.PublishINT('telescope', 'dome', 'POSITION.INSTRUMENTAL.HA.MOTION_STATE', 8);
	ELSE
		fbComm.PublishINT('telescope', 'dome', 'POSITION.INSTRUMENTAL.HA.MOTION_STATE', 1);
	END_IF
ELSE
	fbComm.PublishINT('telescope', 'dome', 'POSITION.INSTRUMENTAL.HA.MOTION_STATE', 0);
END_IF

fbComm.PublishLREAL('telescope', 'dome', 'POSITION.INSTRUMENTAL.HA.CURRPOS', fHourAngleCurrent);
fbComm.PublishLREAL('telescope', 'dome', 'POSITION.INSTRUMENTAL.HA.REALPOS', fHourAngleCurrent-F_HourAngleOffsetOnAxis(fHourAngleOffset, fDeclinationApparent));
fbComm.PublishLREAL('telescope', 'dome', 'POSITION.INSTRUMENTAL.HA.TARGETPOS', fbHourAngle.Position);
fbComm.PublishLREAL('telescope', 'dome', 'POSITION.INSTRUMENTAL.HA.CURRSPEED', fbHourAngle.Velocity);
fbComm.PublishLREAL('telescope', 'dome', 'POSITION.INSTRUMENTAL.HA.TARGETDISTANCE', ABS(fHourAngleCurrent-fbHourAngle.Position));
fbComm.PublishLREAL('telescope', 'dome', 'POSITION.INSTRUMENTAL.HA.OFFSET', fHourAngleOffset);

// > FOCUS
// POWER_STATE
IF fbFocus.Enable THEN
	fbComm.PublishLREAL('telescope', 'dome', 'POSITION.INSTRUMENTAL.FOCUS.POWER_STATE', 1.0);
ELSE
	fbComm.PublishLREAL('telescope', 'dome', 'POSITION.INSTRUMENTAL.FOCUS.POWER_STATE', 0.0);
END_IF
//REFERENCED
IF fbFocus.Calibrated THEN
	fbComm.PublishLREAL('telescope', 'dome', 'POSITION.INSTRUMENTAL.FOCUS.REFERENCED', 1.0);
ELSE
	fbComm.PublishLREAL('telescope', 'dome', 'POSITION.INSTRUMENTAL.FOCUS.REFERENCED', 0.0);
END_IF
//ERROR_STATE
IF fbFocus.Error THEN
	fbComm.PublishINT('telescope', 'dome', 'POSITION.INSTRUMENTAL.FOCUS.ERROR_STATE', fbHourAngle.ErrorID);
ELSE
	fbComm.PublishINT('telescope', 'dome', 'POSITION.INSTRUMENTAL.FOCUS.ERROR_STATE', 0);
END_IF
//MOTION_STATE
IF fbFocus.Busy THEN
	fbComm.PublishINT('telescope', 'dome', 'POSITION.INSTRUMENTAL.FOCUS.MOTION_STATE', 1);
ELSE
	fbComm.PublishINT('telescope', 'dome', 'POSITION.INSTRUMENTAL.FOCUS.MOTION_STATE', 0);
END_IF
fbComm.PublishLREAL('telescope', 'dome', 'POSITION.INSTRUMENTAL.FOCUS.CURRPOS', fbFocus.ActualPosition);
fbComm.PublishLREAL('telescope', 'dome', 'POSITION.INSTRUMENTAL.FOCUS.REALPOS', fbFocus.ActualPosition);
fbComm.PublishLREAL('telescope', 'dome', 'POSITION.INSTRUMENTAL.FOCUS.TARGETPOS', fbFocus.Position);
fbComm.PublishLREAL('telescope', 'dome', 'POSITION.INSTRUMENTAL.FOCUS.TARGETDISTANCE', ABS(fbFocus.ActualPosition-fbFocus.Position));
fbComm.PublishLREAL('telescope', 'dome', 'POSITION.INSTRUMENTAL.FOCUS.CURRSPEED', fbFocus.Velocity);


(*HORIZONTAL*)
fbComm.PublishLREAL('telescope', 'dome', 'POSITION.HORIZONTAL.ALT', fElevationCurrentSky);
fbComm.PublishLREAL('telescope', 'dome', 'POSITION.HORIZONTAL.AZ', fAzimuthCurrentSky);
fbComm.PublishLREAL('telescope', 'dome', 'POSITION.HORIZONTAL.DOME', fbDome.Position);

(*EQUITORIAL*)
fbComm.PublishLREAL('telescope', 'dome', 'POSITION.EQUATORIAL.RA_ICRS', fRightAscensionCurrentICRScorr);	// degrees (BROTLib#37)
fbComm.PublishLREAL('telescope', 'dome', 'POSITION.EQUATORIAL.DEC_ICRS', fDeclinationCurrentICRScorr);
fbComm.PublishLREAL('telescope', 'dome', 'POSITION.EQUATORIAL.HA_APPARENT', fHourAngleCurrent - fHourAngleInversionOffset - F_HourAngleOffsetOnAxis(fHourAngleOffset, fDeclinationApparent));
fbComm.PublishLREAL('telescope', 'dome', 'POSITION.EQUATORIAL.DEC_APPARENT', fDeclinationCurrent - fDeclinationInversionOffset - fDeclinationOffset);
END_METHOD

METHOD PRIVATE _SlewTelescope : USINT
VAR_INPUT
END_VAR
VAR
	SlewEvent:	FB_Eventlog;
END_VAR
VAR_INST
	nStage:		USINT := 0;
	nLastStage:	USINT := 101;
END_VAR
_SlewTelescope := nStage;
IF tonSlewTimeout.Q THEN	// MONETcommon#17: fed every scan in the body
	bSoftwareError := TRUE;		// #30
	nSoftwareErrorID := 16#40;
	bSlewActive := FALSE;
	nStage := 0;
	RETURN;
END_IF
IF bResetActive OR bError OR bStopActive OR bInterrupted THEN
	nStage := 0;
	RETURN;
END_IF
CASE nStage OF
	0:	
		// #42: not gated on bStopped/bTracking any more, stage 10 ends the tracking (like the goto). Waiting for
		// both here hung a slew sent while tracking: the arbitration had already dropped the track command.
		IF bReady AND NOT bBusy THEN
			nStage := 10;
		END_IF
	10:
		IF fbHourAngle.Tracking = TRUE OR fbDeclination.Tracking = TRUE THEN
			fbHourAngle.Tracking := FALSE;
			fbDeclination.Tracking := FALSE;
		ELSE
			nStage := 20;
		END_IF
	20:
		// send Dome position
		THIS^.fbDome.Position := fAzimuth;
		THIS^.HourAngleOffset := 0.0;
		THIS^.DeclinationOffset := 0.0;
		// write the calculated coordinates into the goto coordinates
		THIS^.fDeclination := fDeclinationCalc;
		THIS^.fRightAscension := fRightAscensionCalc;
		nStage := 25;
	25:
		// Declination (including pointing model)
		fbDeclination.Position := fDeclinationCalc + fDeclinationPointingOffset;
		// HourAngle
		// change to -180 to 180 degree in HA
		IF MODABS(fHourangleCalc + fHourAnglePointingOffset, 360) > 180 THEN
			fbHourAngle.Position := MODABS(fHourangleCalc + fHourAnglePointingOffset,360) - 360.0;
		ELSE
			fbHourAngle.Position := MODABS(fHourangleCalc + fHourAnglePointingOffset,360);
		END_IF
		
		fbHourAngle.Velocity := fSlewVelocity;
		fbDeclination.Velocity := fSlewVelocity;
		// make sure to never drive under Horizon
		IF ABS(fbHourAngle.Position) < ABS(fHourangleCalc) THEN
			// move Ha then Dec
			nStage := 30;
		ELSE
			// move Dec then HA
			nStage := 40;
		END_IF
	// Stage 30: move Ha and then Dec
	30:
		fbHourAngle.MoveAxis := TRUE;
		IF fbHourAngle.Busy THEN
			nStage := 31;
		END_IF
	31:
		IF NOT fbHourAngle.Busy AND fbHourAngle.MoveDone THEN
			fbHourAngle.MoveAxis := FALSE;
		END_IF
		IF NOT fbHourAngle.MoveAxis THEN
		   nStage := 32;
		END_IF
	32:
		fbDeclination.MoveAxis := TRUE;
		IF fbDeclination.Busy THEN
			nStage := 33;
		END_IF
	33:
		IF NOT fbDeclination.Busy AND fbDeclination.MoveDone THEN
			fbDeclination.MoveAxis := FALSE;
		END_IF
		IF NOT fbDeclination.MoveAxis THEN
		   nStage := 75;
		END_IF
	// Stage 40: move Dec and then Ha
	40:
		fbDeclination.MoveAxis := TRUE;
		IF fbDeclination.Busy THEN
			nStage := 41;
		END_IF
	41:
		IF NOT fbDeclination.Busy AND fbDeclination.MoveDone THEN
			fbDeclination.MoveAxis := FALSE;
		END_IF
		IF NOT fbDeclination.MoveAxis THEN
		   nStage := 42;
		END_IF
	42:
		fbHourAngle.MoveAxis := TRUE;
		IF fbHourAngle.Busy THEN
			nStage := 43;
		END_IF
	43:
		IF NOT fbHourAngle.Busy AND fbHourAngle.MoveDone THEN
			fbHourAngle.MoveAxis := FALSE;
		END_IF
		IF NOT fbHourAngle.MoveAxis THEN
		   nStage := 75;
		END_IF
	75:
		IF NOT bSliding AND bStopped THEN // all axis standstill
			nStage := 100;
		END_IF
	100:
		fbHourAngle.MoveAxis := FALSE;
		fbDeclination.MoveAxis := FALSE;

		bSlewActive := FALSE;
		nStage := 0;
END_CASE
SlewEvent(Trigger := nStage > nLastStage, FormatString := 'Slew progress: %s', OnMessage := USINT_TO_STRING(nStage), comm := fbComm);
nLastStage := nStage;
END_METHOD

// BROTLib#25 step 4.4a: the inputs of the generic stop transaction (axis 1 = hour angle, 2 = declination), set before the
// body and before Monitor() so that both see this scan's values.
METHOD PRIVATE _SetStopTxInputs
fbStopTx.abEnabled[1] := fbHourAngle.bEnable;
fbStopTx.abEnabled[2] := fbDeclination.bEnable;
fbStopTx.abStandStill[1] := aAxis[1].bStandStill;
fbStopTx.abStandStill[2] := aAxis[2].bStandStill;
fbStopTx.abStopAxis[1] := fbHourAngle.StopAxis;
fbStopTx.abStopAxis[2] := fbDeclination.StopAxis;
fbStopTx.abStopDone[1] := aAxis[1].bStopDone;
fbStopTx.abStopDone[2] := aAxis[2].bStopDone;
fbStopTx.abLocked[1] := (fbHourAngle.axisRef.NcToPlc.StateDWord AND 16#20000000) <> 0;	// MotionCommandsLocked
fbStopTx.abLocked[2] := (fbDeclination.axisRef.NcToPlc.StateDWord AND 16#20000000) <> 0;
fbStopTx.abHoming[1] := fbHourAngle.fbLatchHome.Busy;
fbStopTx.abHoming[2] := fbDeclination.fbLatchHome.Busy;
fbStopTx.abMoving[1] := aAxis[1].bInMotion OR aAxis[1].bInRamp;	// for Restart
fbStopTx.abMoving[2] := aAxis[2].bInMotion OR aAxis[2].bInRamp;
fbStopTx.abStopping[1] := aAxis[1].bStopping;
fbStopTx.abStopping[2] := aAxis[2].bStopping;
fbStopTx.abSweeping[1] := fbHourAngle.bSweepActive;	// #198
fbStopTx.abSweeping[2] := fbDeclination.bSweepActive;
fbStopTx.bStopped := bStopped;
fbStopTx.tTimeout := T#30S;	// #120: the stop command timeout
fbStopTx.nTimeDivisor := nTimeDivisor;
END_METHOD

METHOD PRIVATE _StopTelescope : BOOL
VAR_INPUT
END_VAR
IF fbHourAngle.Tracking = TRUE OR fbDeclination.Tracking = TRUE THEN
	fbHourAngle.Tracking := FALSE;
	fbDeclination.Tracking := FALSE;
ELSIF fbHourAngle.MoveAxis = TRUE OR  fbDeclination.MoveAxis = TRUE THEN
	fbHourAngle.MoveAxis := FALSE;
	fbDeclination.MoveAxis := FALSE;
ELSE
	// Only issue Axis stop commands if they are moving, and only one per axis and stop transaction (#108): a running
	// MC_Stop reports StandStill FALSE, so asking again after every StopDone restarted it about 33 times per second.
	// An axis that finishes a scan later than the other (HA outside its target window after 120 s of tracking) then
	// never lined up with the other one, bStopped stayed FALSE and a gohome waiting for it was dropped. FB_AxisControl
	// clears StopAxis on StopDone.
	_SetStopTxInputs();
	fbStopTx();
	IF fbStopTx.abWriteLow[1] THEN
		fbHourAngle.StopAxis := FALSE;	// a level left TRUE by an earlier stop: low for one scan, the stop follows
	ELSIF fbStopTx.abWriteHigh[1] THEN
		fbHourAngle.StopAxis := TRUE;
	END_IF

	IF fbStopTx.abWriteLow[2] THEN
		fbDeclination.StopAxis := FALSE;
	ELSIF fbStopTx.abWriteHigh[2] THEN
		fbDeclination.StopAxis := TRUE;
	END_IF

	IF fbStopTx.bSettled THEN
		fbHourAngle.StopAxis := FALSE;
		fbDeclination.StopAxis := FALSE;
		_StopTelescope := FALSE;
	END_IF
END_IF
END_METHOD

METHOD PRIVATE _TrackTelescope : BOOL
VAR_INPUT
END_VAR
// send Dome position
THIS^.fbDome.Position := fAzimuthCurrent;
// Declination (including offest and pointing model)
fbDeclination.Position := fDeclinationApparent + fDeclinationOffset + fDeclinationPointingOffset;
// HourAngle
// change to -180 to 180 degree in HA
IF MODABS(fHourAngleApparent + F_HourAngleOffsetOnAxis(fHourAngleOffset, fDeclinationApparent)+ fHourAnglePointingOffset, 360) > 180 THEN
	fbHourAngle.Position := MODABS(fHourAngleApparent + F_HourAngleOffsetOnAxis(fHourAngleOffset, fDeclinationApparent)+ fHourAnglePointingOffset,360) - 360.0;
ELSE
	fbHourAngle.Position := MODABS(fHourAngleApparent + F_HourAngleOffsetOnAxis(fHourAngleOffset, fDeclinationApparent)+ fHourAnglePointingOffset,360);
END_IF


IF NOT fbHourAngle.Tracking THEN
	fbHourAngle.Velocity := 1.0;
	fbHourAngle.MoveAxis := TRUE;
	IF NOT fbHourAngle.Busy AND fbHourAngle.MoveDone THEN
		fbHourAngle.MoveAxis := FALSE;
		IF fbHourAngle.isTracking THEN
			fbHourAngle.Velocity := fHourAngleVelocity;
		END_IF
		fbHourAngle.Tracking := TRUE;
	END_IF
ELSE
	fbHourAngle.Velocity := fHourAngleVelocity;
END_IF


IF NOT fbDeclination.Tracking THEN
	fbDeclination.Velocity := 1.0;
	fbDeclination.MoveAxis := TRUE;
	IF NOT fbDeclination.Busy AND fbDeclination.MoveDone THEN
		fbDeclination.MoveAxis := FALSE;
		IF fbDeclination.isTracking THEN
			fbDeclination.Velocity := fDeclinationVelocity;
		END_IF
		fbDeclination.Tracking := TRUE;
	END_IF
ELSE
	fbDeclination.Velocity := fDeclinationVelocity;
END_IF
END_METHOD

PROPERTY AltAz : BROTLib.ST_AltAzCoordinate
GET
AltAz.Altitude 	:= fElevationCalc;
AltAz.Azimuth 	:= fAzimuthCalc;
END_GET
END_PROPERTY

{warning 'add property implementation'}
PROPERTY Altitude : LREAL
GET
Altitude := fElevationCurrent;
END_GET
END_PROPERTY

{warning 'add property implementation'}
PROPERTY Azimuth : LREAL
GET
Azimuth := fAzimuthCurrent;
END_GET
END_PROPERTY

PROPERTY CoverAutoOpen : BOOL
GET
CoverAutoOpen := bCoverAutoOpen;
END_GET
SET
bCoverAutoOpen := CoverAutoOpen;
END_SET
END_PROPERTY

{warning 'add property implementation'}
PROPERTY Declination : LREAL
GET
END_GET
END_PROPERTY

PROPERTY DeclinationOffset : LREAL
GET
DeclinationOffset := fDeclinationOffset;
END_GET
SET
fDeclinationOffset := DeclinationOffset;
END_SET
END_PROPERTY

//FB_Init is always available implicitly and it is used primarily for initialization.
//The return value is not evaluated. For a specific influence, you can also declare the
//methods explicitly and provide additional code there with the standard initialization
//code. You can evaluate the return value.
METHOD FB_Init: BOOL
VAR_INPUT
    bInitRetains	: BOOL; // TRUE: the retain variables are initialized (reset warm / reset cold)
    bInCopyCode		: BOOL;  // TRUE: the instance will be copied to the copy code afterward (online change)
	comm			: I_Comm;
END_VAR
THIS^.fbComm 				:= comm;
END_METHOD

METHOD Home : BOOL
bGoHomeChecked := TRUE;
// decide first (a home while not ready, powering on or parked is rejected, no longer waited for 2 min); a rejection writes nothing
IF NOT _AcceptMove(E_TCSCommand.gohome, E_TCSCommand.no_command) THEN
	RETURN;
END_IF
bHomeByCommand := TRUE;
bGoHomeActive := TRUE;
Home := TRUE;
END_METHOD

PROPERTY HourAngleOffset : LREAL
GET
HourAngleOffset := fHourAngleOffset;
END_GET
SET
fHourAngleOffset := HourAngleOffset;
END_SET
END_PROPERTY

METHOD Init : BOOL
bPowerChecked := TRUE;
// park wins in both orders and a stop is not overridden by a power-on (MONETcommon#87); this comes before AcceptInit, a pending
// park clears Initialized, so AcceptInit would accept. The in-place park (bSafeParked, up to 120 s) is refused as well.
IF bStopActive OR bParkActive OR bParkAfterStop OR bSafeParked THEN
    nInitRefusedCount := nInitRefusedCount + 1;
    bInitRefused := TRUE;
    IF bStopActive THEN
        sInitRefusedReason := 'stop in progress';
    ELSIF bSafeParked THEN
        sInitRefusedReason := 'in-place park in progress, ends within 120 s';
    ELSE
        sInitRefusedReason := 'park in progress, send stop to cancel it';
    END_IF
// AcceptInit refuses while a startup runs or completed (also across a transient interlock, -2).
ELSIF fbStartup.AcceptInit() THEN
    // nothing stale after the power-on starts: a pending move or home from before would run into it (park is kept, it is the safe direction)
    bGoHomeActive := FALSE;
    bGotoActive := FALSE;
    bSlewActive := FALSE;
    bTrackActive := FALSE;
    bPowerActive := TRUE;
    fReadyState := 0.7;
    // #159: an automatic stop leaves the sweep hold set with the axes enabled; a new power-on releases it
    fbHourAngle.bReleaseHold := TRUE;
    fbDeclination.bReleaseHold := TRUE;
END_IF
Init := TRUE;
END_METHOD

PROPERTY RaDec : BROTLib.ST_RaDecCoordinate
GET
RaDec.RightAscension	:= fRightAscensionCalc;
RaDec.Declination		:= fDeclinationCalc;
END_GET
END_PROPERTY

METHOD Reset : BOOL
bResetChecked := TRUE;
bResetRequest := TRUE;
END_METHOD

// READY_STATE as published on TELESCOPE.READY_STATE; BROTLib.FB_Comm_MQTT_Influx accepts the focus command only at 1 (BROTLib#74)
PROPERTY ReadyState : LREAL
GET
ReadyState := fReadyState;
END_GET
END_PROPERTY

{warning 'add property implementation'}
PROPERTY RightAscension : LREAL
GET
END_GET
END_PROPERTY

METHOD SetAltitudeOffset : BOOL
VAR_INPUT
	Offset	: LREAL;
END_VAR
END_METHOD

METHOD SetAzimuthOffset : BOOL
VAR_INPUT
	Offset	: LREAL;
END_VAR
END_METHOD

METHOD SetDeclinationOffset : BOOL
VAR_INPUT
	Offset	: LREAL;
END_VAR
fDeclinationOffset := Offset;
END_METHOD

METHOD SetDerotatorOffset : BOOL
VAR_INPUT
	Offset	: LREAL;
END_VAR
END_METHOD

METHOD SetRightAscensionOffset : BOOL
VAR_INPUT
	Offset	: LREAL;
END_VAR
fHourAngleOffset := -1.0*Offset;
END_METHOD

{warning 'add method implementation '}
METHOD Slew : BOOL
VAR_INPUT
	fAzimuth	: LREAL;
	fAltitude	: LREAL;
END_VAR
// #100: not while the telescope is not ready (parked, powering on, error). The request used to stay latched and
// fired unnoticed after the next power-on; a client sends init first and waits for ready.
bSlewChecked := TRUE;
// decided at arrival (F_CommandAcceptance): a rejected slew writes nothing, not even the target, and is never left pending
IF NOT _AcceptMove(E_TCSCommand.slew, E_TCSCommand.no_command) THEN
	RETURN;
END_IF
THIS^.fElevation 	:= fAltitude;
THIS^.fAzimuth 	:= fAzimuth;
bSlewActive		:= TRUE;
END_METHOD

METHOD Stop : BOOL
bStopChecked := TRUE;
// a stop ends a park that is queued behind a running stop (MONETcommon#213)
bParkAfterStop := FALSE;
// a repeated stop while a stop is running sends a new stop only to axes that are moving again and are not stopping already
// (BROTLib.FB_StopTransaction.Restart); the focus is stopped again as well (MONETcommon#96/#122)
IF bStopActive THEN
	_SetStopTxInputs();
	fbStopTx.Restart();
	IF fbFocus <> 0 THEN
		fbFocus.Stop();
	END_IF
END_IF
bStopActive := TRUE;
// MONETcommon#122: an explicit stop also stops a running focus move and holds the position reached; the automatic
// stops of the mount (horizon, pole zone) leave the focus alone
IF fbFocus <> 0 THEN
	fbFocus.Stop();
END_IF
END_METHOD

{warning 'add method implementation '}
METHOD Track : BOOL
VAR_INPUT
	fRightAscension	: LREAL;
	fDeclination	: LREAL;
END_VAR
// #100: see Slew(); a track request while the telescope is not ready is refused, not latched
bGotoChecked := TRUE;
bTrackChecked := TRUE;	// D4 (template body step S1.f): Track() and a bTrack edge in one scan are one command, as in MONETcommon
IF NOT _AcceptMove(E_TCSCommand.goto, E_TCSCommand.no_command) THEN
	RETURN;
END_IF
THIS^.fRightAscension	:= fRightAscension;
THIS^.fDeclination	:= fDeclination;
bGotoActive			:= TRUE;
END_METHOD

END_FUNCTION_BLOCK

// ---- POUs/FB_CabinetControl.TcPOU
FUNCTION_BLOCK FB_CabinetControl
VAR_INPUT
	bEstop				: BOOL;	// E-stop pressed (telescope bEstopTriggered, previous scan) (#93)
	bSafetyAckPending	: BOOL;	// safety acknowledge after an E-stop not yet run, drives still in STO (#93)
END_VAR
VAR_OUTPUT
END_VAR
VAR
	bCabinetError : BOOL;
	bTelescopeError : BOOL;
	bReset	: BOOL;
	
	rtrigReset : R_TRIG;
	
	bAuxiliaryContact24V AT %I* : BOOL; // Auxilary Contact of the 24V DC: TRUE = operational
	bAuxiliaryContact48V AT %I* : BOOL; // Auxilary Contact of the 48V DC: TRUE = operational
	bAuxiliaryContactHADEC AT %I* : BOOL; // Auxilary Contact of the HA DEC motor: TRUE = operational
	bAuxiliaryContactFOCUS AT %I* : BOOL; // Auxilary Contact of the FOCUS motor: TRUE = operational
	bCollectiveReport24VFuse AT %I*: BOOL; // Collective Report of the 24V Fuse box: TRUE = operational
	bState24VFuse AT %I*: BOOL; 
	
	bOErrorLED	AT %Q* : BOOL;
	bIReset     AT %I* : BOOL;
	bIMode      AT %I* : BOOL;
END_VAR

// #10: error when ANY of the five is lost (it was NOT(a OR b OR ...), which only fired when all five dropped).
// All five read TRUE parked, powered and at three E-stops (test T14, 2026-10-12/13), so none of them is FALSE in
// normal operation. bState24VFuse is FALSE throughout and stays out of the expression.
bCabinetError := NOT( bAuxiliaryContact24V AND bAuxiliaryContact48V AND bAuxiliaryContactHADEC AND bAuxiliaryContactFOCUS AND bCollectiveReport24VFuse);

// if error -> LED on
// #93: also while the E-stop is pressed and until the safety acknowledge has run (the drives are in STO and a reset
// is needed). Not part of bError, which would change the reset condition, the power-on block and STATUS.GLOBAL.
bOErrorLED := bTelescopeError OR bEstop OR bSafetyAckPending;

// if reset -> trigger reset
rtrigReset(CLK:= bIReset,Q=>bReset);

PROPERTY Error : BOOL
GET
Error := bCabinetError;
END_GET
SET
bTelescopeError := Error;
END_SET
END_PROPERTY

PROPERTY LocalMode : BOOL
GET
LocalMode := bIMode;
END_GET
END_PROPERTY

PROPERTY Reset : BOOL
GET
Reset := bReset;
END_GET
END_PROPERTY

END_FUNCTION_BLOCK

// ---- POUs/Pointing/FB_PointingModelForward.TcPOU
FUNCTION_BLOCK FB_PointingModelForward
VAR_INPUT
	HourAngle		: LREAL;
	Declination		: LREAL;
	Latitude		: LREAL;
END_VAR
VAR_OUTPUT
	HourAngle_correction	: LREAL;
	Declination_correction	: LREAL;
	HourAngle_velocity		: LREAL;
	Declination_velocity 	: LREAL; 
END_VAR
VAR
	// inputs in rad
	tau		: LREAL;
	dec		: LREAL;
	alt		: LREAL;
	lat		: LREAL;
	// offsets
	off_tau_esti : LREAL :=0.0;
	off_dec_esti : LREAL :=0.0;
	// trackingspeeds
	track_tau_esti : LREAL := 0.0;
	track_dec_esti : LREAL := 0.0;
	// Altitude
	alt_diff : LREAL;
	// pre calculated sin/cos
	sin_tau	: LREAL;
	cos_tau	: LREAL;
	sin_dec	: LREAL;
	cos_dec : LREAL;
	sin_lat	: LREAL;
	cos_lat : LREAL;
	sin_alt : LREAL;
	sin_alt_rate : LREAL;
	cos_alt : LREAL;
END_VAR
VAR CONSTANT
	d2r		: LREAL := PI/180.0;
	omega 	: LREAL := 360.0 / 86164.099 * (PI/180.0); //sidereal velocity
END_VAR

// degrees to rad
tau := HourAngle * d2r;
dec	:= Declination * d2r;
lat := Latitude * d2r;


// pre-calculate repeating sine and cosine functions
sin_TAU := SIN(tau);
cos_TAU := COS(tau);
sin_DEC := SIN(dec);
cos_DEC := COS(dec);
sin_lat := SIN(lat);
cos_lat := COS(lat);

// alt difference estimation (WITHOUT Nutation, Aberation, Presession)
sin_alt := sin_DEC * sin_lat + cos_DEC * cos_lat * cos_TAU;
sin_alt := LIMIT(-1.0, sin_alt, 1.0);	// rounding can give 1 + 2.2E-16 at the zenith, ASIN of that is NaN (#4)
alt := ASIN(sin_alt);					// diagnostics only, not used below
cos_alt := SQRT(1.0 - sin_alt * sin_alt);	// = COS(alt) >= 0
// d(sin alt)/dt = cos(alt) * d(alt)/dt. Finite everywhere; d(alt)/dt itself is 0/0 at the zenith (#4)
sin_alt_rate := -omega * cos_DEC * cos_lat * sin_TAU;
IF cos_alt > 1.0E-9 THEN
	alt_diff := sin_alt_rate / cos_alt;	// diagnostics only, not used below
ELSE
	alt_diff := 0.0;
END_IF

// ### TAU offset ###
off_tau_esti := - C_mAl_tau * ((cos_TAU * sin_DEC) / cos_DEC);
off_tau_esti := off_tau_esti + C_mEl_tau * ((sin_TAU * sin_DEC) / cos_DEC);
off_tau_esti := off_tau_esti + C_Coll_tau;
off_tau_esti := off_tau_esti + C_Refr_tau * ((sin_TAU * cos_lat) / (sin_alt * cos_DEC)); 
off_tau_esti := off_tau_esti + C_Flex_tau * ((sin_TAU * cos_lat) / cos_DEC);
off_tau_esti := off_tau_esti + C_Enc_tau / cos_DEC;
off_tau_esti := off_tau_esti - C_NP_tau * (sin_DEC / cos_DEC);


track_tau_esti := c_mal_tau * omega * ((sin_TAU * sin_DEC) / cos_DEC);
track_tau_esti := track_tau_esti + c_mel_tau * omega * ((cos_TAU * sin_DEC) / cos_DEC);
track_tau_esti := track_tau_esti + c_refr_tau * omega * ((cos_TAU * cos_lat) / (sin_alt * cos_DEC)); // 1ST derivative term
track_tau_esti := track_tau_esti - c_refr_tau * sin_alt_rate * ((sin_TAU * cos_lat) / (sin_alt*sin_alt * cos_DEC)); // 2nd term
track_tau_esti := track_tau_esti + c_flex_tau * omega * ((cos_TAU * cos_lat) / cos_DEC);


// ### DEC offset ###
off_dec_esti := C_mAl_dec * sin_TAU;
off_dec_esti := off_dec_esti + C_mEl_dec * cos_TAU;
off_dec_esti := off_dec_esti + C_Coll_dec;
off_dec_esti := off_dec_esti + C_Refr_dec * ((sin_lat - sin_alt * sin_DEC) / (cos_DEC * sin_alt));
off_dec_esti := off_dec_esti - C_Flex_dec * ((sin_lat - sin_alt * sin_DEC) / cos_DEC);


track_dec_esti := c_mal_dec * omega * cos_TAU;
track_dec_esti := track_dec_esti - c_mel_dec * omega * sin_TAU;
track_dec_esti := track_dec_esti - c_refr_dec * sin_alt_rate * (sin_DEC / (cos_DEC * sin_alt));//# 1ST term
track_dec_esti := track_dec_esti - c_refr_dec * sin_alt_rate * ((sin_lat - sin_alt * sin_DEC) / (cos_DEC * sin_alt*sin_alt)); //# 2nd derivative term
track_dec_esti := track_dec_esti + c_flex_dec * sin_alt_rate * (sin_DEC / cos_DEC);

HourAngle_correction	:= off_tau_esti;
Declination_correction	:= off_dec_esti;
HourAngle_velocity		:= (track_tau_esti + omega)/d2r;
Declination_velocity 	:= track_dec_esti/d2r;

END_FUNCTION_BLOCK

// ---- POUs/Pointing/FB_PointingModelInversion.TcPOU
FUNCTION_BLOCK FB_PointingModelInversion
VAR_INPUT
	HourAngle		: LREAL;
	Declination		: LREAL;
	Altitude		: LREAL;
	Latitude		: LREAL;
	epsilon			: LREAL := 0.25; //iteration accuracy in arcsec
END_VAR
VAR_OUTPUT
	HourAngle_correction	: LREAL;
	Declination_correction	: LREAL;
	bValid					: BOOL;	// FALSE if the iteration did not converge within epsilon (e.g. altitude too close to the horizon, where the model is chaotic -- see testing/check_pointing_inversion.py). HourAngle_correction/Declination_correction are 0.0 when FALSE.
END_VAR
VAR
	fbpointing : FB_PointingModelForward;
	d_ha		: LREAL := 0.0;
	d_dec		: LREAL := 0.0;
	d_ha_new	: LREAL := 0.0;
	d_dec_new	: LREAL := 0.0;
	i			: INT;
	
END_VAR

